      #   Source: Robotiq_Grippers, 1.8.4.4844, Robotiq Inc.
      #   Type: Gripper
      $ 2003 "Gripper Close (1)"
      if not(gripper_connected[0]):
        popup("Gripper 1 must be connected to run this program.", "No connection", False, True, True)
      end
      if not(rq_is_gripper_activated("1")):
        popup("Gripper 1 is not activated. Go to Installation tab > Gripper to activate it and run the program again.", "Not activated", False, True, True)
      end
      rq_set_pos_spd_for(255, 204, 255, "1")
      rq_wait_pos_spe_for_request(255, 204, 255, "1")
      rq_go_to("1")
      rq_wait("1")
      # end: URCap Program Node
      $ 2010 "Decap"
      $ 2011 "Action_Info≔'decapping'"
      global Action_Info="decapping"
      $ 2012 "Set GRP_3F_Enable=On"
      set_standard_digital_out(4, True)
      $ 2013 "Set GRP_3F_Decap=On"
      set_standard_digital_out(3, True)
      $ 2014 "Force"
      sleep(0.02)
      zero_ftsensor()
      force_mode(p[0.0,0.0,0.0,0.0,0.0,0.0], [0, 0, 1, 0, 0, 0], [0.0, 0.0, 1.0, 0.0, 0.0, 0.0], 2, [0.1, 0.1, 0.001, 0.3490658503988659, 0.3490658503988659, 0.3490658503988659])
      $ 2015 "check_decapping(offset=0.015, timeout=10, abort=CMD_Hold)" "noBreak"
      check_decapping(offset=0.015, timeout=10, abort=CMD_Hold)
      end_force_mode()
      stopl(5.0)
      $ 2016 "Set GRP_3F_Decap=Off"
      set_standard_digital_out(3, False)
      $ 2017 "Set GRP_3F_Enable=Off"
      set_standard_digital_out(4, False)
      $ 2018 "MoveL"
      $ 2019 "Waypoint_50" "breakAfter"
      movel(Waypoint_50_p, a=0.5, v=0.1, r=0.05)
      $ 2020 "MoveJ"
      $ 2021 "cap_dump" "breakAfter"
      movej(get_inverse_kin(cap_dump_p, qnear=cap_dump_q), a=0.5235987755982988, v=0.4363323129985824)
      # begin: URCap Program Node
      #   Source: Robotiq_Grippers, 1.8.4.4844, Robotiq Inc.
      #   Type: Gripper
      $ 2022 "Gripper Open (1)"
      if not(gripper_connected[0]):
        popup("Gripper 1 must be connected to run this program.", "No connection", False, True, True)
      end
      if not(rq_is_gripper_activated("1")):
        popup("Gripper 1 is not activated. Go to Installation tab > Gripper to activate it and run the program again.", "Not activated", False, True, True)
      end
      rq_set_pos_spd_for(0, 204, 255, "1")
      rq_wait_pos_spe_for_request(0, 204, 255, "1")
      rq_go_to("1")
      rq_wait("1")
      # end: URCap Program Node
      $ 2023 "MoveJ"
      $ 2024 "Waypoint_51" "breakAfter"
      movej(get_inverse_kin(Waypoint_51_p, qnear=Waypoint_51_q), a=0.5235987755982988, v=0.4363323129985824, r=0.036)
    elif (33 == switch_1):
      $ 2025 "Case 33"
      $ 2026 "Shake and liquid transfer"
      $ 2027 "MoveL"
      $ 2028 "Vial_liq_above" "breakAfter"
      movel(Vial_liq_above_p, a=0.5, v=0.1)
      $ 2029 "Vial_liq_pick_1" "breakAfter"
      movel(Vial_liq_pick_1_p, a=0.5, v=0.1)
      $ 2030 "Vial_liq_pick_2" "breakAfter"
      movel(Vial_liq_pick_2_p, a=0.5, v=0.1)
      # begin: URCap Program Node
      #   Source: Robotiq_Grippers, 1.8.4.4844, Robotiq Inc.
      #   Type: Gripper
      $ 2031 "Gripper Close (1)"
      if not(gripper_connected[0]):
        popup("Gripper 1 must be connected to run this program.", "No connection", False, True, True)
      end
      if not(rq_is_gripper_activated("1")):
        popup("Gripper 1 is not activated. Go to Installation tab > Gripper to activate it and run the program again.", "Not activated", False, True, True)
      end
      rq_set_pos_spd_for(255, 82, 71, "1")
      rq_wait_pos_spe_for_request(255, 82, 71, "1")
      rq_go_to("1")
      rq_wait("1")
      # end: URCap Program Node
      $ 2032 "Wait: 1.0"
      sleep(1.0)
      $ 2033 "Set GRP_3F_Open=On"
      set_standard_digital_out(5, True)
      $ 2034 "Wait: 0.5"
      sleep(0.5)
      $ 2035 "Vial_liq_above" "breakAfter"
      movel(Vial_liq_above_p, a=0.3, v=0.05, r=0.05)
      $ 2036 "MoveL"
      $ 2037 "Liquid_midway" "breakAfter"
      movel(Liquid_midway_p, a=0.5, v=0.1)
      $ 2038 "Loop 3 times"
      Loop_1 = 0
      while (Loop_1 < 3):
        $ 2039 "shake_1" "breakAfter"
        movel(shake_1_p, a=2.0, v=0.5)
        $ 2040 "shake_2" "breakAfter"
        movel(shake_2_p, a=2.0, v=0.5)
        Loop_1 = Loop_1 + 1
      end
      $ 2041 "drop_above_1" "breakAfter"
      movel(drop_above_1_p, a=0.5, v=0.1)
      $ 2042 "drop_above_2" "breakAfter"
      movel(drop_above_2_p, a=0.5, v=0.1)
      $ 2043 "liq_tran_1" "breakAfter"
      movel(liq_tran_1_p, a=0.5, v=0.05, r=0.008)
      $ 2044 "Wait: 1.0"
      sleep(1.0)
      $ 2045 "drop_above_2" "breakAfter"
      movel(drop_above_2_p, a=0.5, v=0.1)
      $ 2046 "Waypoint_21" "breakAfter"
      movel(Waypoint_21_p, a=0.5, v=0.1)
      $ 2047 "liq_tran_2" "breakAfter"
      movel(liq_tran_2_p, a=0.5, v=0.05)
      $ 2048 "Wait: 1.0"
      sleep(1.0)
      $ 2049 "drop_above_2" "breakAfter"
      movel(drop_above_2_p, a=0.5, v=0.1)
      $ 2050 "drop_above_1" "breakAfter"
      movel(drop_above_1_p, a=0.5, v=0.1)
      $ 2051 "Liquid_midway" "breakAfter"
      movel(Liquid_midway_p, a=0.5, v=0.1)
      $ 2052 "MoveL"
      $ 2053 "Vial_drop_above" "breakAfter"
      movel(Vial_drop_above_p, a=0.5, v=0.1)
      $ 2054 "Vial_liq_drop" "breakAfter"
      movel(Vial_liq_drop_p, a=0.5, v=0.1)
      # begin: URCap Program Node
      #   Source: Robotiq_Grippers, 1.8.4.4844, Robotiq Inc.
      #   Type: Gripper
      $ 2055 "Gripper Open (1)"
      if not(gripper_connected[0]):
        popup("Gripper 1 must be connected to run this program.", "No connection", False, True, True)
      end
      if not(rq_is_gripper_activated("1")):
        popup("Gripper 1 is not activated. Go to Installation tab > Gripper to activate it and run the program again.", "Not activated", False, True, True)
      end
      rq_set_pos_spd_for(0, 82, 71, "1")
      rq_wait_pos_spe_for_request(0, 82, 71, "1")
      rq_go_to("1")
      rq_wait("1")
      # end: URCap Program Node
      $ 2056 "Vial_drop_above" "breakAfter"
      movel(Vial_drop_above_p, a=0.5, v=0.1)
    elif (34 == switch_1):
      $ 2057 "Case 34"
      $ 2058 "Home (Safe)"
      movej([-1.2302089344500047, -1.2969853503591224, -1.875639182904262, -1.539621866126728, 1.5731943360401213, -2.80099559440227], a=1.3962634015954636, v=1.0471975511965976)
      $ 2059 "MoveJ"
      $ 2060 "Waypoint_9" "breakAfter"
      movej(get_inverse_kin(Waypoint_9_p, qnear=Waypoint_9_q), a=0.5235987755982988, v=0.4363323129985824)
      $ 2061 "MoveL"
      $ 2062 "Waypoint_10" "breakAfter"
      movel(Waypoint_10_p, a=0.5, v=0.1)
      # begin: URCap Program Node
      #   Source: Robotiq_Grippers, 1.8.4.4844, Robotiq Inc.
      #   Type: Gripper
      $ 2063 "Gripper Close (1)"
      if not(gripper_connected[0]):
        popup("Gripper 1 must be connected to run this program.", "No connection", False, True, True)
      end
      if not(rq_is_gripper_activated("1")):
        popup("Gripper 1 is not activated. Go to Installation tab > Gripper to activate it and run the program again.", "Not activated", False, True, True)
      end
      rq_set_pos_spd_for(255, 82, 71, "1")
      rq_wait_pos_spe_for_request(255, 82, 71, "1")
      rq_go_to("1")
      rq_wait("1")
      # end: URCap Program Node
      $ 2064 "Wait: 1.0"
      sleep(1.0)
      $ 2065 "MoveL"
      $ 2066 "Waypoint_11" "breakAfter"
      movel(Waypoint_11_p, a=0.5, v=0.1, r=0.05)
      $ 2067 "MoveJ"
      $ 2068 "Waypoint_7" "breakAfter"
      movej(get_inverse_kin(Waypoint_7_p, qnear=Waypoint_7_q), a=0.5235987755982988, v=0.4363323129985824, r=0.05)
      $ 2069 "MoveL"
      $ 2070 "Waypoint_8" "breakAfter"
      movel(Waypoint_8_p, a=0.5, v=0.1)
      # begin: URCap Program Node
      #   Source: Robotiq_Grippers, 1.8.4.4844, Robotiq Inc.
      #   Type: Gripper
      $ 2071 "Gripper Open (1)"
      if not(gripper_connected[0]):
        popup("Gripper 1 must be connected to run this program.", "No connection", False, True, True)
      end
      if not(rq_is_gripper_activated("1")):
        popup("Gripper 1 is not activated. Go to Installation tab > Gripper to activate it and run the program again.", "Not activated", False, True, True)
      end
      rq_set_pos_spd_for(0, 82, 71, "1")
      rq_wait_pos_spe_for_request(0, 82, 71, "1")
      rq_go_to("1")
      rq_wait("1")
      # end: URCap Program Node
      $ 2072 "MoveJ"
      $ 2073 "Waypoint_7" "breakAfter"
      movej(get_inverse_kin(Waypoint_7_p, qnear=Waypoint_7_q), a=0.5235987755982988, v=0.4363323129985824)
      $ 2074 "Home (Safe)"
      movej([-1.2302089344500047, -1.2969853503591224, -1.875639182904262, -1.539621866126728, 1.5731943360401213, -2.80099559440227], a=1.3962634015954636, v=1.0471975511965976)
    elif (35 == switch_1):
      $ 2091 "Case 35"
      $ 2092 "Pick the powder container"
      $ 2093 "Wait: 1.0"
      sleep(1.0)
      $ 2094 "MoveJ"
      $ 2095 "Container_midwa" "breakAfter"
      movej(get_inverse_kin(Container_midwa_p, qnear=Container_midwa_q), a=1.3962634015954636, v=1.0471975511965976, r=0.05)
      $ 2096 "Container_capt" "breakAfter"
      movej(get_inverse_kin(Container_capt_p, qnear=Container_capt_q), a=1.3962634015954636, v=1.0471975511965976)
      # begin: URCap Program Node
      #   Source: SensoPart VISOR Robotic, 2.0.0, SensoPart Industriesensorik GmbH
      #   Type: VISOR Robotic App
      $ 2097 "VISOR Easy Pick"
      def visorFuncEasyPick_e3134b():
        # begin: URCap Program Node
        #   Source: SensoPart VISOR Robotic, 2.0.0, SensoPart Industriesensorik GmbH
        #   Type: Easy Pick Setup
        $ 2098 "# 1 Setup" "noBreak"
        local easyPickVisorId = 1
        local easyPickArmMounted = True
        local easyPickSetJob = True
        local easyPickJobName = "Container_S"
        local easyPickAtImgAcq = False
        local easyPickImgAcqPose = p[-0.5104,0.4173,0.4641,0.0000,-0.0000,-2.8962]
        # end: URCap Program Node
        # begin: URCap Program Node
        #   Source: SensoPart VISOR Robotic, 2.0.0, SensoPart Industriesensorik GmbH
        #   Type: Process
        $ 2099 "Process" "noBreak"
        local easyPickObjTaken = False
        local easyPickTrigger = False
        local easyPickPoseIdx = 0
        local easyPickPose = p[0,0,0,0,0,0]
        def easyPickFuncTrigger(visorId, setJob, jobName, arm):
        if (setJob):
          visor_changeJob(visorId, jobName, 6000)
        end
        if (arm):
          visor_trigger(visorId, 6000, "arm")
        else:
          visor_trigger(visorId, 6000)
        end
        global easyPickParts=visor_partsFound(visorId)
        visor_easyPickUpdate(visorId, "parts", visor_partsFound(visorId))
        return visor_getPose3d(visorId, 0)
      end
      while (not easyPickObjTaken):
        easyPickTrigger = (easyPickCount >= visor_partsFound(easyPickVisorId)) or (easyPickCount > 9) or (not visor_easyPickCheckIdent("70ff7e", easyPickVisorId))
        if (easyPickTrigger):
          easyPickCount = 0
        end
        easyPickPoseIdx = easyPickCount
        easyPickPose = visor_getPose3d(easyPickVisorId, easyPickPoseIdx)
        visor_easyPickUpdate(easyPickVisorId, "counter", easyPickPoseIdx)
        # begin: URCap Program Node
        #   Source: SensoPart VISOR Robotic, 2.0.0, SensoPart Industriesensorik GmbH
        #   Type: Image Acquisition Pose
        $ 2100 "Image Acquisition Pose" "noBreak"
        if (easyPickTrigger):
          if (not easyPickAtImgAcq):
            movej(pose_trans(easyPickImgAcqPose,p[0.0000,0.0000,-0.0000,0.0000,0.0000,0.0000]),a=1.3963,v=1.0472,t=0.000000,r=0.000000)
            easyPickAtImgAcq = True
          end
          easyPickPose = easyPickFuncTrigger(easyPickVisorId, easyPickSetJob, easyPickJobName, easyPickArmMounted)
        end
        # end: URCap Program Node
        # begin: URCap Program Node
        #   Source: SensoPart VISOR Robotic, 2.0.0, SensoPart Industriesensorik GmbH
        #   Type: Object Detected
        $ 2101 "Object Detected" "noBreak"
        if (visor_partsFound(easyPickVisorId) > 0):
          $ 2102 "Open Gripper" "noBreak"
          # begin: URCap Program Node
          #   Source: Robotiq_Grippers, 1.8.4.4844, Robotiq Inc.
          #   Type: Gripper
          $ 2103 "Gripper Open (1)" "noBreak"
          if not(gripper_connected[0]):
            popup("Gripper 1 must be connected to run this program.", "No connection", False, True, True)
          end
          if not(rq_is_gripper_activated("1")):
            popup("Gripper 1 is not activated. Go to Installation tab > Gripper to activate it and run the program again.", "Not activated", False, True, True)
          end
          rq_set_pos_spd_for(0, 107, 77, "1")
          rq_wait_pos_spe_for_request(0, 107, 77, "1")
          rq_go_to("1")
          rq_wait("1")
          # end: URCap Program Node
          $ 2104 "MoveJ" "noBreak"
          $ 2105 "Waypoint_13" "noBreak"
          movej(get_inverse_kin(Waypoint_13_p, qnear=Waypoint_13_q), a=1.3962634015954636, v=1.0471975511965976)
          # begin: URCap Program Node
          #   Source: SensoPart VISOR Robotic, 2.0.0, SensoPart Industriesensorik GmbH
          #   Type: Approach Pose
          $ 2106 "Approach Pose" "noBreak"
          movej(pose_trans(easyPickPose,p[0.0000,0.0000,0.0500,0.0000,0.0000,0.0000]),a=1.3963,v=1.0472,t=0.000000,r=0.000000)
          # end: URCap Program Node
          # begin: URCap Program Node
          #   Source: SensoPart VISOR Robotic, 2.0.0, SensoPart Industriesensorik GmbH
          #   Type: Target Pose
          $ 2107 "Target Pose" "noBreak"
          movel(pose_trans(easyPickPose,p[0.0000,0.0000,-0.0000,0.0000,0.0000,0.0000]),a=0.5000,v=0.2500,t=0.000000,r=0.000000)
          # end: URCap Program Node
          $ 2108 "Close Gripper" "noBreak"
          # begin: URCap Program Node
          #   Source: Robotiq_Grippers, 1.8.4.4844, Robotiq Inc.
          #   Type: Gripper
          $ 2109 "Gripper Close (1)" "noBreak"
          if not(gripper_connected[0]):
            popup("Gripper 1 must be connected to run this program.", "No connection", False, True, True)
          end
          if not(rq_is_gripper_activated("1")):
            popup("Gripper 1 is not activated. Go to Installation tab > Gripper to activate it and run the program again.", "Not activated", False, True, True)
          end
          rq_set_pos_spd_for(255, 107, 77, "1")
          rq_wait_pos_spe_for_request(255, 107, 77, "1")
          rq_go_to("1")
          rq_wait("1")
          # end: URCap Program Node
          # begin: URCap Program Node
          #   Source: SensoPart VISOR Robotic, 2.0.0, SensoPart Industriesensorik GmbH
          #   Type: Exit Pose
          $ 2110 "Exit Pose" "noBreak"
          movel(pose_trans(easyPickPose,p[0.0000,0.0000,0.0500,0.0000,0.0000,0.0000]),a=0.5000,v=0.2500,t=0.000000,r=0.000000)
          # end: URCap Program Node
          easyPickObjTaken = True
        end
        # end: URCap Program Node
        # begin: URCap Program Node
        #   Source: SensoPart VISOR Robotic, 2.0.0, SensoPart Industriesensorik GmbH
        #   Type: No Object Detected
        $ 2111 "No Object Detected" "noBreak"
        if (visor_partsFound(easyPickVisorId) < 1):
          easyPickNoObj = easyPickNoObj + 1
          if (easyPickNoObj > 5):
            global easyPickNoObj=0
            halt
          end
          $ 2112 "Popup: No Container detected" "noBreak"
          popup("No Container detected", "Message", False, False, blocking=True)
          else:
          global easyPickNoObj=0
        end
        # end: URCap Program Node
      end
      easyPickCount = easyPickCount + 1
      visor_easyPickUpdate(easyPickVisorId, "counter", easyPickCount)
      visor_easyPickSetIdent("70ff7e", easyPickVisorId)
      # end: URCap Program Node
    end
    visorFuncEasyPick_e3134b()
    # end: URCap Program Node
    $ 2113 "MoveJ"
    $ 2114 "Cont_midwa_1" "breakAfter"
    movej(get_inverse_kin(Cont_midwa_1_p, qnear=Cont_midwa_1_q), a=1.3962634015954636, v=1.0471975511965976, r=0.05)
    $ 2115 "Cont_midw_2" "breakAfter"
    movej(get_inverse_kin(Cont_midw_2_p, qnear=Cont_midw_2_q), a=1.3962634015954636, v=1.0471975511965976, r=0.05)
    $ 2116 "MoveJ"
    $ 2117 "Waypoint_14" "breakAfter"
    movej(get_inverse_kin(Waypoint_14_p, qnear=Waypoint_14_q), a=1.3962634015954636, v=1.0471975511965976)
    $ 2118 "Cont_midway_3" "breakAfter"
    movej(get_inverse_kin(Cont_midway_3_p, qnear=Cont_midway_3_q), a=1.3962634015954636, v=1.0471975511965976)
    $ 2119 "Waypoint_43" "breakAfter"
    movej(get_inverse_kin(Waypoint_43_p, qnear=Waypoint_43_q), a=1.3962634015954636, v=1.0471975511965976)
    $ 2120 "MoveL"
    $ 2121 "Waypoint_27" "breakAfter"
    movel(Waypoint_27_p, a=1.2, v=0.25)
    $ 2122 "Waypoint_2" "breakAfter"
    movel(Waypoint_2_p, a=0.3, v=0.05)
    # begin: URCap Program Node
    #   Source: Robotiq_Grippers, 1.8.4.4844, Robotiq Inc.
    #   Type: Gripper
    $ 2123 "Gripper Open (1)"
    if not(gripper_connected[0]):
      popup("Gripper 1 must be connected to run this program.", "No connection", False, True, True)
    end
    if not(rq_is_gripper_activated("1")):
      popup("Gripper 1 is not activated. Go to Installation tab > Gripper to activate it and run the program again.", "Not activated", False, True, True)
    end
    rq_set_pos_spd_for(0, 255, 255, "1")
    rq_wait_pos_spe_for_request(0, 255, 255, "1")
    rq_go_to("1")
    rq_wait("1")
    # end: URCap Program Node
    $ 2124 "MoveL"
    $ 2125 "Waypoint_27" "breakAfter"
    movel(Waypoint_27_p, a=1.2, v=0.25)
    $ 2126 "Waypoint_39" "breakAfter"
    movel(Waypoint_39_p, a=1.2, v=0.25)
    $ 2127 "Home (Safe)"
    movej([-1.2302089344500047, -1.2969853503591224, -1.875639182904262, -1.539621866126728, 1.5731943360401213, -2.80099559440227], a=1.3962634015954636, v=1.0471975511965976)
    # begin: URCap Program Node
    #   Source: SensoPart VISOR Robotic, 2.0.0, SensoPart Industriesensorik GmbH
    #   Type: VISOR Robotic App
    $ 2128 "VISOR Easy Pick"
    def visorFuncEasyPick_ffc504():
      # begin: URCap Program Node
      #   Source: SensoPart VISOR Robotic, 2.0.0, SensoPart Industriesensorik GmbH
      #   Type: Easy Pick Setup
      $ 2129 "# 1 Setup" "noBreak"
      local easyPickVisorId = 1
      local easyPickArmMounted = True
      local easyPickSetJob = True
      local easyPickJobName = "Target_container"
      local easyPickAtImgAcq = False
      local easyPickImgAcqPose = p[-0.6180,0.3719,0.4116,-0.0000,-0.0000,-2.8962]
      # end: URCap Program Node
      # begin: URCap Program Node
      #   Source: SensoPart VISOR Robotic, 2.0.0, SensoPart Industriesensorik GmbH
      #   Type: Process
      $ 2130 "Process" "noBreak"
      local easyPickObjTaken = False
      local easyPickTrigger = False
      local easyPickPoseIdx = 0
      local easyPickPose = p[0,0,0,0,0,0]
      def easyPickFuncTrigger(visorId, setJob, jobName, arm):
      if (setJob):
        visor_changeJob(visorId, jobName, 6000)
      end
      if (arm):
        visor_trigger(visorId, 6000, "arm")
      else:
        visor_trigger(visorId, 6000)
      end
      global easyPickParts_2=visor_partsFound(visorId)
      visor_easyPickUpdate(visorId, "parts", visor_partsFound(visorId))
      return visor_getPose3d(visorId, 0)
    end
    while (not easyPickObjTaken):
      easyPickTrigger = (easyPickCount_2 >= visor_partsFound(easyPickVisorId)) or (easyPickCount_2 > 9) or (not visor_easyPickCheckIdent("9ee82b", easyPickVisorId))
      if (easyPickTrigger):
        easyPickCount_2 = 0
      end
      easyPickPoseIdx = easyPickCount_2
      easyPickPose = visor_getPose3d(easyPickVisorId, easyPickPoseIdx)
      visor_easyPickUpdate(easyPickVisorId, "counter", easyPickPoseIdx)
      # begin: URCap Program Node
      #   Source: SensoPart VISOR Robotic, 2.0.0, SensoPart Industriesensorik GmbH
      #   Type: Image Acquisition Pose
      $ 2131 "Image Acquisition Pose" "noBreak"
      if (easyPickTrigger):
        if (not easyPickAtImgAcq):
          movej(pose_trans(easyPickImgAcqPose,p[0.0000,0.0000,-0.0000,0.0000,0.0000,0.0000]),a=1.3963,v=1.0472,t=0.000000,r=0.000000)
          easyPickAtImgAcq = True
        end
        easyPickPose = easyPickFuncTrigger(easyPickVisorId, easyPickSetJob, easyPickJobName, easyPickArmMounted)
      end
      # end: URCap Program Node
      # begin: URCap Program Node
      #   Source: SensoPart VISOR Robotic, 2.0.0, SensoPart Industriesensorik GmbH
      #   Type: Object Detected
      $ 2132 "Object Detected" "noBreak"
      if (visor_partsFound(easyPickVisorId) > 0):
        $ 2133 "Open Gripper" "noBreak"
        # begin: URCap Program Node
        #   Source: Robotiq_Grippers, 1.8.4.4844, Robotiq Inc.
        #   Type: Gripper
        $ 2134 "Gripper Open (1)" "noBreak"
        if not(gripper_connected[0]):
          popup("Gripper 1 must be connected to run this program.", "No connection", False, True, True)
        end
        if not(rq_is_gripper_activated("1")):
          popup("Gripper 1 is not activated. Go to Installation tab > Gripper to activate it and run the program again.", "Not activated", False, True, True)
        end
        rq_set_pos_spd_for(0, 107, 77, "1")
        rq_wait_pos_spe_for_request(0, 107, 77, "1")
        rq_go_to("1")
        rq_wait("1")
        # end: URCap Program Node
        # begin: URCap Program Node
        #   Source: SensoPart VISOR Robotic, 2.0.0, SensoPart Industriesensorik GmbH
        #   Type: Approach Pose
        $ 2135 "Approach Pose" "noBreak"
        movej(pose_trans(easyPickPose,p[0.0000,0.0000,0.0500,0.0000,0.0000,0.0000]),a=1.3963,v=1.0472,t=0.000000,r=0.000000)
        # end: URCap Program Node
        # begin: URCap Program Node
        #   Source: SensoPart VISOR Robotic, 2.0.0, SensoPart Industriesensorik GmbH
        #   Type: Target Pose
        $ 2136 "Target Pose" "noBreak"
        movel(pose_trans(easyPickPose,p[0.0000,0.0000,-0.0000,0.0000,0.0000,0.0000]),a=0.5000,v=0.2500,t=0.000000,r=0.000000)
        # end: URCap Program Node
        $ 2137 "Close Gripper" "noBreak"
        # begin: URCap Program Node
        #   Source: Robotiq_Grippers, 1.8.4.4844, Robotiq Inc.
        #   Type: Gripper
        $ 2138 "Gripper Close (1)" "noBreak"
        if not(gripper_connected[0]):
          popup("Gripper 1 must be connected to run this program.", "No connection", False, True, True)
        end
        if not(rq_is_gripper_activated("1")):
          popup("Gripper 1 is not activated. Go to Installation tab > Gripper to activate it and run the program again.", "Not activated", False, True, True)
        end
        rq_set_pos_spd_for(255, 107, 77, "1")
        rq_wait_pos_spe_for_request(255, 107, 77, "1")
        rq_go_to("1")
        rq_wait("1")
        # end: URCap Program Node
        # begin: URCap Program Node
        #   Source: SensoPart VISOR Robotic, 2.0.0, SensoPart Industriesensorik GmbH
        #   Type: Exit Pose
        $ 2139 "Exit Pose" "noBreak"
        movel(pose_trans(easyPickPose,p[0.0000,0.0000,0.0500,0.0000,0.0000,0.0000]),a=0.5000,v=0.2500,t=0.000000,r=0.000000)
        # end: URCap Program Node
        easyPickObjTaken = True
      end
      # end: URCap Program Node
      # begin: URCap Program Node
      #   Source: SensoPart VISOR Robotic, 2.0.0, SensoPart Industriesensorik GmbH
      #   Type: No Object Detected
      $ 2140 "No Object Detected" "noBreak"
      if (visor_partsFound(easyPickVisorId) < 1):
        easyPickNoObj_2 = easyPickNoObj_2 + 1
        if (easyPickNoObj_2 > 5):
          global easyPickNoObj_2=0
          halt
        end
        $ 2141 "Popup: No target container is detected" "noBreak"
        popup("No target container is detected", "Message", False, False, blocking=True)
        else:
        global easyPickNoObj_2=0
      end
      # end: URCap Program Node
    end
    easyPickCount_2 = easyPickCount_2 + 1
    visor_easyPickUpdate(easyPickVisorId, "counter", easyPickCount_2)
    visor_easyPickSetIdent("9ee82b", easyPickVisorId)
    # end: URCap Program Node
  end
  visorFuncEasyPick_ffc504()
  # end: URCap Program Node
  $ 2142 "MoveJ"
  $ 2143 "Waypoint_5" "breakAfter"
  movej(get_inverse_kin(Waypoint_5_p, qnear=Waypoint_5_q), a=1.3962634015954636, v=1.0471975511965976)
  $ 2144 "Waypoint_3" "breakAfter"
  movej(get_inverse_kin(Waypoint_3_p, qnear=Waypoint_3_q), a=1.3962634015954636, v=1.0471975511965976)
  $ 2145 "Set GRP_3F_Open=On"
  set_standard_digital_out(5, True)
  $ 2146 "MoveL"
  $ 2147 "Waypoint_4" "breakAfter"
  movel(Waypoint_4_p, a=1.2, v=0.25)
  $ 2148 "Waypoint_15" "breakAfter"
  movel(Waypoint_15_p, a=0.3, v=0.05)
  $ 2149 "Set GRP_3F_Open=Off"
  set_standard_digital_out(5, False)
  $ 2150 "Wait: 0.5"
  sleep(0.5)
  # begin: URCap Program Node
  #   Source: Robotiq_Grippers, 1.8.4.4844, Robotiq Inc.
  #   Type: Gripper
  $ 2151 "Gripper Open (1)"
  if not(gripper_connected[0]):
    popup("Gripper 1 must be connected to run this program.", "No connection", False, True, True)
  end
  if not(rq_is_gripper_activated("1")):
    popup("Gripper 1 is not activated. Go to Installation tab > Gripper to activate it and run the program again.", "Not activated", False, True, True)
  end
  rq_set_pos_spd_for(0, 127, 71, "1")
  rq_wait_pos_spe_for_request(0, 127, 71, "1")
  rq_go_to("1")
  rq_wait("1")
  # end: URCap Program Node
  $ 2152 "MoveL"
  $ 2153 "Waypoint_16" "breakAfter"
  movel(Waypoint_16_p, a=1.2, v=0.25)
  $ 2154 "Home (Safe)"
  movej([-1.2302089344500047, -1.2969853503591224, -1.875639182904262, -1.539621866126728, 1.5731943360401213, -2.80099559440227], a=1.3962634015954636, v=1.0471975511965976)
  elif (36 == switch_1):
    $ 2155 "Case 36"
    $ 2156 "MoveJ"
    $ 2157 "Waypoint_23" "breakAfter"
    movej(get_inverse_kin(Waypoint_23_p, qnear=Waypoint_23_q), a=1.3962634015954636, v=1.0471975511965976)
    $ 2158 "MoveL"
    $ 2159 "Waypoint_24" "breakAfter"
    movel(Waypoint_24_p, a=1.2, v=0.25)
    # begin: URCap Program Node
    #   Source: Robotiq_Grippers, 1.8.4.4844, Robotiq Inc.
    #   Type: Gripper
    $ 2160 "Gripper Close (1)"
    if not(gripper_connected[0]):
      popup("Gripper 1 must be connected to run this program.", "No connection", False, True, True)
    end
    if not(rq_is_gripper_activated("1")):
      popup("Gripper 1 is not activated. Go to Installation tab > Gripper to activate it and run the program again.", "Not activated", False, True, True)
    end
    rq_set_pos_spd_for(255, 127, 127, "1")
    rq_wait_pos_spe_for_request(255, 127, 127, "1")
    rq_go_to("1")
    rq_wait("1")
    # end: URCap Program Node
    $ 2161 "Decap"
    $ 2162 "Action_Info≔'decapping'"
    global Action_Info="decapping"
    $ 2163 "Set GRP_3F_Enable=On"
    set_standard_digital_out(4, True)
    $ 2164 "Set GRP_3F_Decap=On"
    set_standard_digital_out(3, True)
    $ 2165 "Force"
    sleep(0.02)
    zero_ftsensor()
    force_mode(p[0.0,0.0,0.0,0.0,0.0,0.0], [0, 0, 1, 0, 0, 0], [0.0, 0.0, 1.0, 0.0, 0.0, 0.0], 2, [0.1, 0.1, 0.001, 0.3490658503988659, 0.3490658503988659, 0.3490658503988659])
    $ 2166 "check_decapping(offset=0.08, timeout=16, abort=CMD_Hold)" "noBreak"
    check_decapping(offset=0.08, timeout=16, abort=CMD_Hold)
    end_force_mode()
    stopl(5.0)
    $ 2167 "Set GRP_3F_Decap=Off"
    set_standard_digital_out(3, False)
    $ 2168 "Set GRP_3F_Enable=Off"
    set_standard_digital_out(4, False)
    $ 2169 "MoveL"
    $ 2170 "Waypoint_17" "breakAfter"
    movel(Waypoint_17_p, a=1.2, v=0.25)
    $ 2171 "Waypoint_22" "breakAfter"
    movel(Waypoint_22_p, a=1.2, v=0.25)
    $ 2172 "Waypoint_25" "breakAfter"
    movel(Waypoint_25_p, a=1.2, v=0.25)
    # begin: URCap Program Node
    #   Source: Robotiq_Grippers, 1.8.4.4844, Robotiq Inc.
    #   Type: Gripper
    $ 2173 "Gripper Open (1)"
    if not(gripper_connected[0]):
      popup("Gripper 1 must be connected to run this program.", "No connection", False, True, True)
    end
    if not(rq_is_gripper_activated("1")):
      popup("Gripper 1 is not activated. Go to Installation tab > Gripper to activate it and run the program again.", "Not activated", False, True, True)
    end
    rq_set_pos_spd_for(0, 107, 77, "1")
    rq_wait_pos_spe_for_request(0, 107, 77, "1")
    rq_go_to("1")
    rq_wait("1")
    # end: URCap Program Node
    $ 2174 "MoveL"
    $ 2175 "Waypoint_26" "breakAfter"
    movel(Waypoint_26_p, a=1.2, v=0.25)
    $ 2176 "MoveL"
    $ 2177 "Waypoint_30" "breakAfter"
    movel(Waypoint_30_p, a=1.2, v=0.25)
    $ 2178 "Waypoint_28" "breakAfter"
    movel(Waypoint_28_p, a=1.2, v=0.25)
    # begin: URCap Program Node
    #   Source: Robotiq_Grippers, 1.8.4.4844, Robotiq Inc.
    #   Type: Gripper
    $ 2179 "Gripper Close (1)"
    if not(gripper_connected[0]):
      popup("Gripper 1 must be connected to run this program.", "No connection", False, True, True)
    end
    if not(rq_is_gripper_activated("1")):
      popup("Gripper 1 is not activated. Go to Installation tab > Gripper to activate it and run the program again.", "Not activated", False, True, True)
    end
    rq_set_pos_spd_for(255, 107, 77, "1")
    rq_wait_pos_spe_for_request(255, 107, 77, "1")
    rq_go_to("1")
    rq_wait("1")
    # end: URCap Program Node
    $ 2180 "Wait: 0.5"
    sleep(0.5)
    $ 2181 "Set GRP_3F_Open=On"
    set_standard_digital_out(5, True)
    $ 2182 "MoveL"
    $ 2183 "Waypoint_29" "breakAfter"
    movel(Waypoint_29_p, a=1.2, v=0.25)
    $ 2184 "MoveJ"
    $ 2185 "Waypoint_31" "breakAfter"
    movej(get_inverse_kin(Waypoint_31_p, qnear=Waypoint_31_q), a=1.3962634015954636, v=1.0471975511965976)
    # begin: URCap Program Node
    #   Source: SensoPart VISOR Robotic, 2.0.0, SensoPart Industriesensorik GmbH
    #   Type: VISOR Robotic App
    $ 2186 "VISOR Easy Pick"
    def visorFuncEasyPick_7a8a4a():
      # begin: URCap Program Node
      #   Source: SensoPart VISOR Robotic, 2.0.0, SensoPart Industriesensorik GmbH
      #   Type: Easy Pick Setup
      $ 2187 "# 1 Setup" "noBreak"
      local easyPickVisorId = 1
      local easyPickArmMounted = True
      local easyPickSetJob = True
      local easyPickJobName = "Weigh_scale"
      local easyPickAtImgAcq = False
      local easyPickImgAcqPose = p[-0.6121,0.0166,0.5300,0.0440,-0.0067,-1.6589]
      # end: URCap Program Node
      # begin: URCap Program Node
      #   Source: SensoPart VISOR Robotic, 2.0.0, SensoPart Industriesensorik GmbH
      #   Type: Process
      $ 2188 "Process" "noBreak"
      local easyPickObjTaken = False
      local easyPickTrigger = False
      local easyPickPoseIdx = 0
      local easyPickPose = p[0,0,0,0,0,0]
      def easyPickFuncTrigger(visorId, setJob, jobName, arm):
      if (setJob):
        visor_changeJob(visorId, jobName, 6000)
      end
      if (arm):
        visor_trigger(visorId, 6000, "arm")
      else:
        visor_trigger(visorId, 6000)
      end
      global easyPickParts_1=visor_partsFound(visorId)
      visor_easyPickUpdate(visorId, "parts", visor_partsFound(visorId))
      return visor_getPose3d(visorId, 0)
    end
    while (not easyPickObjTaken):
      easyPickTrigger = (easyPickCount_1 >= visor_partsFound(easyPickVisorId)) or (easyPickCount_1 > 9) or (not visor_easyPickCheckIdent("425780", easyPickVisorId))
      if (easyPickTrigger):
        easyPickCount_1 = 0
      end
      easyPickPoseIdx = easyPickCount_1
      easyPickPose = visor_getPose3d(easyPickVisorId, easyPickPoseIdx)
      visor_easyPickUpdate(easyPickVisorId, "counter", easyPickPoseIdx)
      # begin: URCap Program Node
      #   Source: SensoPart VISOR Robotic, 2.0.0, SensoPart Industriesensorik GmbH
      #   Type: Image Acquisition Pose
      $ 2189 "Image Acquisition Pose" "noBreak"
      if (easyPickTrigger):
        if (not easyPickAtImgAcq):
          movej(pose_trans(easyPickImgAcqPose,p[0.0000,0.0000,-0.0000,0.0000,0.0000,0.0000]),a=1.3963,v=1.0472,t=0.000000,r=0.000000)
          easyPickAtImgAcq = True
        end
        easyPickPose = easyPickFuncTrigger(easyPickVisorId, easyPickSetJob, easyPickJobName, easyPickArmMounted)
      end
      # end: URCap Program Node
      # begin: URCap Program Node
      #   Source: SensoPart VISOR Robotic, 2.0.0, SensoPart Industriesensorik GmbH
      #   Type: Object Detected
      $ 2190 "Object Detected" "noBreak"
      if (visor_partsFound(easyPickVisorId) > 0):
        $ 2191 "Open Gripper" "noBreak"
        $ 2192 "Wait: 0.5" "noBreak"
        sleep(0.5)
        # begin: URCap Program Node
        #   Source: SensoPart VISOR Robotic, 2.0.0, SensoPart Industriesensorik GmbH
        #   Type: Approach Pose
        $ 2193 "Approach Pose" "noBreak"
        movej(pose_trans(easyPickPose,p[0.0000,0.0000,0.0300,0.0000,0.0000,0.0000]),a=1.3963,v=1.0472,t=0.000000,r=0.000000)
        # end: URCap Program Node
        # begin: URCap Program Node
        #   Source: SensoPart VISOR Robotic, 2.0.0, SensoPart Industriesensorik GmbH
        #   Type: Target Pose
        $ 2194 "Target Pose" "noBreak"
        movel(pose_trans(easyPickPose,p[0.0000,0.0000,-0.0000,0.0000,0.0000,0.0000]),a=0.5000,v=0.2500,t=0.000000,r=0.000000)
        # end: URCap Program Node
        $ 2195 "Close Gripper" "noBreak"
        # begin: URCap Program Node
        #   Source: Robotiq_Grippers, 1.8.4.4844, Robotiq Inc.
        #   Type: Gripper
        $ 2196 "Gripper Open (1)" "noBreak"
        if not(gripper_connected[0]):
          popup("Gripper 1 must be connected to run this program.", "No connection", False, True, True)
        end
        if not(rq_is_gripper_activated("1")):
          popup("Gripper 1 is not activated. Go to Installation tab > Gripper to activate it and run the program again.", "Not activated", False, True, True)
        end
        rq_set_pos_spd_for(0, 255, 255, "1")
        rq_wait_pos_spe_for_request(0, 255, 255, "1")
        rq_go_to("1")
        rq_wait("1")
        # end: URCap Program Node
        # begin: URCap Program Node
        #   Source: SensoPart VISOR Robotic, 2.0.0, SensoPart Industriesensorik GmbH
        #   Type: Exit Pose
        $ 2197 "Exit Pose" "noBreak"
        movel(pose_trans(easyPickPose,p[0.0000,0.0000,0.0500,0.0000,0.0000,0.0000]),a=0.5000,v=0.2500,t=0.000000,r=0.000000)
        # end: URCap Program Node
        easyPickObjTaken = True
      end
      # end: URCap Program Node
      # begin: URCap Program Node
      #   Source: SensoPart VISOR Robotic, 2.0.0, SensoPart Industriesensorik GmbH
      #   Type: No Object Detected
      $ 2198 "No Object Detected" "noBreak"
      if (visor_partsFound(easyPickVisorId) < 1):
        $ 2199 "Popup: No weigh scale detected" "noBreak"
        popup("No weigh scale detected", "Message", False, False, blocking=True)
        else:
      end
      # end: URCap Program Node
    end
    easyPickCount_1 = easyPickCount_1 + 1
    visor_easyPickUpdate(easyPickVisorId, "counter", easyPickCount_1)
    visor_easyPickSetIdent("425780", easyPickVisorId)
    # end: URCap Program Node
  end
  visorFuncEasyPick_7a8a4a()
  # end: URCap Program Node
  $ 2200 "MoveJ"
  $ 2201 "Waypoint_46" "breakAfter"
  movej(get_inverse_kin(Waypoint_46_p, qnear=Waypoint_46_q), a=1.3962634015954636, v=1.0471975511965976, r=0.05)
  $ 2202 "Waypoint_32" "breakAfter"
  movej(get_inverse_kin(Waypoint_32_p, qnear=Waypoint_32_q), a=1.3962634015954636, v=1.0471975511965976, r=0.011)
  $ 2203 "MoveL"
  $ 2204 "Waypoint_33" "breakAfter"
  movel(Waypoint_33_p, a=1.2, v=0.25, r=0.05)
  $ 2205 "Waypoint_34" "breakAfter"
  movel(Waypoint_34_p, a=1.2, v=0.25, r=0.009000000000000001)
  # begin: URCap Program Node
  #   Source: Robotiq_Grippers, 1.8.4.4844, Robotiq Inc.
  #   Type: Gripper
  $ 2206 "Gripper Move10mm (1)"
  if not(gripper_connected[0]):
    popup("Gripper 1 must be connected to run this program.", "No connection", False, True, True)
  end
  if not(rq_is_gripper_activated("1")):
    popup("Gripper 1 is not activated. Go to Installation tab > Gripper to activate it and run the program again.", "Not activated", False, True, True)
  end
  rq_set_pos_spd_for(203, 64, 62, "1")
  rq_wait_pos_spe_for_request(203, 64, 62, "1")
  rq_go_to("1")
  rq_wait("1")
  # end: URCap Program Node
  $ 2207 "MoveL"
  $ 2208 "Waypoint_40" "breakAfter"
  movel(Waypoint_40_p, a=1.2, v=0.25, r=0.001)
  $ 2209 "decap_1" "breakAfter"
  movel(decap_1_p, a=1.2, v=0.25)
  # begin: URCap Program Node
  #   Source: Robotiq_Grippers, 1.8.4.4844, Robotiq Inc.
  #   Type: Gripper
  $ 2210 "Gripper Move45mm (1)"
  if not(gripper_connected[0]):
    popup("Gripper 1 must be connected to run this program.", "No connection", False, True, True)
  end
  if not(rq_is_gripper_activated("1")):
    popup("Gripper 1 is not activated. Go to Installation tab > Gripper to activate it and run the program again.", "Not activated", False, True, True)
  end
  rq_set_pos_spd_for(40, 173, 153, "1")
  rq_wait_pos_spe_for_request(40, 173, 153, "1")
  rq_go_to("1")
  rq_wait("1")
  # end: URCap Program Node
  $ 2211 "MoveL"
  $ 2212 "Waypoint_41" "breakAfter"
  movel(Waypoint_41_p, a=1.2, v=0.25)
  $ 2213 "Waypoint_42" "breakAfter"
  movel(Waypoint_42_p, a=1.2, v=0.25)
  $ 2214 "decap_2" "breakAfter"
  movel(decap_2_p, a=1.2, v=0.25)
  # begin: URCap Program Node
  #   Source: Robotiq_Grippers, 1.8.4.4844, Robotiq Inc.
  #   Type: Gripper
  $ 2215 "Gripper Move10mm (1)"
  if not(gripper_connected[0]):
    popup("Gripper 1 must be connected to run this program.", "No connection", False, True, True)
  end
  if not(rq_is_gripper_activated("1")):
    popup("Gripper 1 is not activated. Go to Installation tab > Gripper to activate it and run the program again.", "Not activated", False, True, True)
  end
  rq_set_pos_spd_for(203, 99, 79, "1")
  rq_wait_pos_spe_for_request(203, 99, 79, "1")
  rq_go_to("1")
  rq_wait("1")
  # end: URCap Program Node
  $ 2216 "MoveL"
  $ 2217 "Waypoint_44" "breakAfter"
  movel(Waypoint_44_p, a=1.2, v=0.25)
  $ 2218 "Waypoint_45" "breakAfter"
  movel(Waypoint_45_p, a=1.2, v=0.25)
  $ 2219 "decap_1" "breakAfter"
  movel(decap_1_p, a=1.2, v=0.25)
  $ 2220 "Waypoint_35" "breakAfter"
  movel(Waypoint_35_p, a=1.2, v=0.25)
  $ 2221 "Waypoint_36" "breakAfter"
  movel(Waypoint_36_p, a=1.2, v=0.25)
  $ 2222 "Waypoint_37" "breakAfter"
  movel(Waypoint_37_p, a=1.2, v=0.25, r=0.05)
  $ 2223 "Waypoint_38" "breakAfter"
  movel(Waypoint_38_p, a=1.2, v=0.25, r=0.05)
  # begin: URCap Program Node
  #   Source: Robotiq_Grippers, 1.8.4.4844, Robotiq Inc.
  #   Type: Gripper
  $ 2224 "Gripper Move38mm (1)"
  if not(gripper_connected[0]):
    popup("Gripper 1 must be connected to run this program.", "No connection", False, True, True)
  end
  if not(rq_is_gripper_activated("1")):
    popup("Gripper 1 is not activated. Go to Installation tab > Gripper to activate it and run the program again.", "Not activated", False, True, True)
  end
  rq_set_pos_spd_for(73, 173, 153, "1")
  rq_wait_pos_spe_for_request(73, 173, 153, "1")
  rq_go_to("1")
  rq_wait("1")
  # end: URCap Program Node
  $ 2225 "MoveL"
  $ 2226 "Waypoint_37" "breakAfter"
  movel(Waypoint_37_p, a=1.2, v=0.25, r=0.05)
  $ 2227 "Home (Safe)"
  movej([-1.2302089344500047, -1.2969853503591224, -1.875639182904262, -1.539621866126728, 1.5731943360401213, -2.80099559440227], a=1.3962634015954636, v=1.0471975511965976)
  elif (37 == switch_1):
    $ 2228 "Case 37"
    $ 2229 "Detect spatula and powder transfer"
    # begin: URCap Program Node
    #   Source: SensoPart VISOR Robotic, 2.0.0, SensoPart Industriesensorik GmbH
    #   Type: VISOR Robotic App
    $ 2230 "VISOR Easy Pick"
    def visorFuncEasyPick_ff889b():
      # begin: URCap Program Node
      #   Source: SensoPart VISOR Robotic, 2.0.0, SensoPart Industriesensorik GmbH
      #   Type: Easy Pick Setup
      $ 2231 "# 1 Setup" "noBreak"
      local easyPickVisorId = 1
      local easyPickArmMounted = True
      local easyPickSetJob = True
      local easyPickJobName = "Spatula"
      local easyPickAtImgAcq = False
      local easyPickImgAcqPose = p[-0.1334,-0.4212,0.2049,-0.9203,1.0979,-1.4781]
      # end: URCap Program Node
      # begin: URCap Program Node
      #   Source: SensoPart VISOR Robotic, 2.0.0, SensoPart Industriesensorik GmbH
      #   Type: Process
      $ 2232 "Process" "noBreak"
      local easyPickObjTaken = False
      local easyPickTrigger = False
      local easyPickPoseIdx = 0
      local easyPickPose = p[0,0,0,0,0,0]
      def easyPickFuncTrigger(visorId, setJob, jobName, arm):
      if (setJob):
        visor_changeJob(visorId, jobName, 6000)
      end
      if (arm):
        visor_trigger(visorId, 6000, "arm")
      else:
        visor_trigger(visorId, 6000)
      end
      global easyPickParts_3=visor_partsFound(visorId)
      visor_easyPickUpdate(visorId, "parts", visor_partsFound(visorId))
      return visor_getPose3d(visorId, 0)
    end
    while (not easyPickObjTaken):
      easyPickTrigger = (easyPickCount_3 >= visor_partsFound(easyPickVisorId)) or (easyPickCount_3 > 9) or (not visor_easyPickCheckIdent("edc17a", easyPickVisorId))
      if (easyPickTrigger):
        easyPickCount_3 = 0
      end
      easyPickPoseIdx = easyPickCount_3
      easyPickPose = visor_getPose3d(easyPickVisorId, easyPickPoseIdx)
      visor_easyPickUpdate(easyPickVisorId, "counter", easyPickPoseIdx)
      # begin: URCap Program Node
      #   Source: SensoPart VISOR Robotic, 2.0.0, SensoPart Industriesensorik GmbH
      #   Type: Image Acquisition Pose
      $ 2233 "Image Acquisition Pose" "noBreak"
      if (easyPickTrigger):
        if (not easyPickAtImgAcq):
          movej(pose_trans(easyPickImgAcqPose,p[0.0000,0.0000,-0.0000,0.0000,0.0000,0.0000]),a=1.3963,v=1.0472,t=0.000000,r=0.000000)
          easyPickAtImgAcq = True
        end
        easyPickPose = easyPickFuncTrigger(easyPickVisorId, easyPickSetJob, easyPickJobName, easyPickArmMounted)
      end
      # end: URCap Program Node
      # begin: URCap Program Node
      #   Source: SensoPart VISOR Robotic, 2.0.0, SensoPart Industriesensorik GmbH
      #   Type: Object Detected
      $ 2234 "Object Detected" "noBreak"
      if (visor_partsFound(easyPickVisorId) > 0):
        $ 2235 "Open Gripper" "noBreak"
        # begin: URCap Program Node
        #   Source: Robotiq_Grippers, 1.8.4.4844, Robotiq Inc.
        #   Type: Gripper
        $ 2236 "Gripper Open (1)" "noBreak"
        if not(gripper_connected[0]):
          popup("Gripper 1 must be connected to run this program.", "No connection", False, True, True)
        end
        if not(rq_is_gripper_activated("1")):
          popup("Gripper 1 is not activated. Go to Installation tab > Gripper to activate it and run the program again.", "Not activated", False, True, True)
        end
        rq_set_pos_spd_for(0, 130, 89, "1")
        rq_wait_pos_spe_for_request(0, 130, 89, "1")
        rq_go_to("1")
        rq_wait("1")
        # end: URCap Program Node
        # begin: URCap Program Node
        #   Source: SensoPart VISOR Robotic, 2.0.0, SensoPart Industriesensorik GmbH
        #   Type: Approach Pose
        $ 2237 "Approach Pose" "noBreak"
        movej(pose_trans(easyPickPose,p[0.0000,0.0000,0.1000,0.0000,0.0000,0.0000]),a=1.3963,v=1.0472,t=0.000000,r=0.000000)
        # end: URCap Program Node
        # begin: URCap Program Node
        #   Source: SensoPart VISOR Robotic, 2.0.0, SensoPart Industriesensorik GmbH
        #   Type: Target Pose
        $ 2238 "Target Pose" "noBreak"
        movel(pose_trans(easyPickPose,p[0.0000,0.0000,-0.0000,0.0000,0.0000,0.0000]),a=0.5000,v=0.2500,t=0.000000,r=0.000000)
        # end: URCap Program Node
        $ 2239 "Close Gripper" "noBreak"
        # begin: URCap Program Node
        #   Source: Robotiq_Grippers, 1.8.4.4844, Robotiq Inc.
        #   Type: Gripper
        $ 2240 "Gripper Close (1)" "noBreak"
        if not(gripper_connected[0]):
          popup("Gripper 1 must be connected to run this program.", "No connection", False, True, True)
        end
        if not(rq_is_gripper_activated("1")):
          popup("Gripper 1 is not activated. Go to Installation tab > Gripper to activate it and run the program again.", "Not activated", False, True, True)
        end
        rq_set_pos_spd_for(255, 130, 89, "1")
        rq_wait_pos_spe_for_request(255, 130, 89, "1")
        rq_go_to("1")
        rq_wait("1")
        # end: URCap Program Node
        # begin: URCap Program Node
        #   Source: SensoPart VISOR Robotic, 2.0.0, SensoPart Industriesensorik GmbH
        #   Type: Exit Pose
        $ 2241 "Exit Pose" "noBreak"
        movel(pose_trans(easyPickPose,p[0.0000,0.0000,0.2000,0.0000,0.0000,0.0000]),a=0.5000,v=0.2500,t=0.000000,r=0.000000)
        # end: URCap Program Node
        easyPickObjTaken = True
      end
      # end: URCap Program Node
      # begin: URCap Program Node
      #   Source: SensoPart VISOR Robotic, 2.0.0, SensoPart Industriesensorik GmbH
      #   Type: No Object Detected
      $ 2242 "No Object Detected" "noBreak"
      if (visor_partsFound(easyPickVisorId) < 1):
        $ 2243 "Popup: No spatula is detected" "noBreak"
        popup("No spatula is detected", "Message", False, False, blocking=True)
        else:
      end
      # end: URCap Program Node
    end
    easyPickCount_3 = easyPickCount_3 + 1
    visor_easyPickUpdate(easyPickVisorId, "counter", easyPickCount_3)
    visor_easyPickSetIdent("edc17a", easyPickVisorId)
    # end: URCap Program Node
  end
  visorFuncEasyPick_ff889b()
  # end: URCap Program Node
  $ 2244 "MoveL"
  $ 2245 "Waypoint_52" "breakAfter"
  movel(Waypoint_52_p, a=1.2, v=0.25)
  $ 2246 "Waypoint_53" "breakAfter"
  movel(Waypoint_53_p, a=0.3, v=0.05)
  $ 2247 "Loop 2 times"
  Loop_2 = 0
  while (Loop_2 < 2):
    $ 2248 "Waypoint_54" "breakAfter"
    global move_thread_flag_2248=0
    thread move_thread_2248():
      enter_critical
      move_thread_flag_2248 = 1
      movel(Waypoint_54_p, a=0.3, v=0.05)
      move_thread_flag_2248 = 2
      exit_critical
    end
    move_thread_flag_2248 = 0
    move_thread_han_2248 = run move_thread_2248()
    while (True):
      local targetTcpDirection=get_target_tcp_speed()
      local stepsToRetract=tool_contact(direction=targetTcpDirection)
      if (stepsToRetract > 0):
        kill move_thread_han_2248
        stopl(3.0)
        local backTrackMovement=get_actual_joint_positions_history(stepsToRetract)
        local contactPose=get_forward_kin(backTrackMovement)
        local posDir=[targetTcpDirection[0],targetTcpDirection[1],targetTcpDirection[2]]
        local retractTo=contactPose
        if (norm(posDir) > 1e-6):
          local normalizedPosDir=normalize(posDir)
          local additionalRetraction=p[normalizedPosDir[0] * 0.0, normalizedPosDir[1] * 0.0, normalizedPosDir[2] * 0.0, 0, 0, 0]
          retractTo = pose_sub(contactPose, additionalRetraction)
        end
        movel(retractTo, a=3.0, v=0.1)
        $ 2249 "Until (tool_contact_detection)"
        break
      end
      sleep(1.0E-10)
      if (move_thread_flag_2248 > 1):
        join move_thread_han_2248
        break
      end
      sync()
    end
    $ 2250 "Waypoint_55" "breakAfter"
    movel(Waypoint_55_p, a=0.3, v=0.05)
    $ 2251 "Waypoint_56" "breakAfter"
    movel(Waypoint_56_p, a=0.3, v=0.05)
    Loop_2 = Loop_2 + 1
  end
  $ 2252 "Waypoint_57" "breakAfter"
  movel(Waypoint_57_p, a=1.5, v=0.75)
  $ 2253 "Waypoint_56" "breakAfter"
  movel(Waypoint_56_p, a=0.3, v=0.05, r=0.016999999999999998)
  $ 2254 "Waypoint_58" "breakAfter"
  movel(Waypoint_58_p, a=0.3, v=0.05, r=0.05)
  $ 2255 "Waypoint_59" "breakAfter"
  movel(Waypoint_59_p, a=0.3, v=0.05, r=0.05)
  $ 2256 "Waypoint_60" "breakAfter"
  movel(Waypoint_60_p, a=1.2, v=0.25, r=0.05)
  $ 2257 "Waypoint_61" "breakAfter"
  movel(Waypoint_61_p, a=1.2, v=0.25, r=0.05)
  $ 2258 "Waypoint_62" "breakAfter"
  movel(Waypoint_62_p, a=1.2, v=0.25)
  $ 2259 "Waypoint_63" "breakAfter"
  global move_thread_flag_2259=0
  thread move_thread_2259():
    enter_critical
    move_thread_flag_2259 = 1
    movel(Waypoint_63_p, a=0.1, v=0.02)
    move_thread_flag_2259 = 2
    exit_critical
  end
  move_thread_flag_2259 = 0
  move_thread_han_2259 = run move_thread_2259()
  while (True):
    sleep(1.0E-10)
    if (move_thread_flag_2259 > 1):
      join move_thread_han_2259
      break
    end
    sync()
  end
  end
  $ 2278 "'=========='"
  # '=========='
  $ 2279 "PostSettings"
  $ 2280 "'ADD ADDITIONAL CHECKS'"
  # 'ADD ADDITIONAL CHECKS'
  end
  $ 2 "BeforeStart"
  $ 3 "Scripts"
  $ 4 "Script: 001 SCRIPT Errors and Warnings Deifnes V0.2.script"

  #*****************************************************
  # customer          :   UK Essen
  # project name      :   P1132
  #****************************************************
  # controller        :
  # software          :
  #****************************************************
  # author            :   E.Petrichenko
  # Copyright (c)     :   United Robotics Group Health and Food GmbH
  #                       An der Riede 2
  #                       28816 Stuhr
  #                       Germany
  #****************************************************
  # description       :   centrifuge actions for the application
  # version:      	:   0.1
  # created           :   22.08.2024
  # updated           :
  #****************************************************
  # modifications     :
  #
  # date              :
  # name              :
  # reason            :
  #****************************************************


  #################################### VARIABLES DEFINITIONS ###################################

  ERROR_POSE_NOT_REACHABLE = 1002
  ERROR_ROBOT_ARM_NOT_IN_HOME_POSE = 1006
  ERROR_NO_OBJECT_TO_PICK = 1010
  ERROR_NOT_DOCKED = 2003
  ERROR_NOT_REACHABLE_TARGET = 2007
  ERROR_CHARGING_NOT_STARTED = 2008
  ERROR_AMR_WRONG_MODE = 2009
  ERROR_UNKNOWN_POSE = 2010
  ERROR_NO_LANDMARK = 3002
  ERROR_WRONG_ORDER = 4002
  ERROR_CENTRIFUGE_CONNECTION = 5001
  ERROR_CENTRIFUGE_POWER = 5002
  ERROR_CENTRIFUGE = 5003
  ERROR_CENTRIFUGE_LID = 5004
  ERROR_CANNOT_OPEN_HATCH = 5006
  ERROR_CANNOT_CLOSE_HATCH = 5008
  ERROR_CANNOT_ROTATE = 5010
  ERROR_CANNOT_START = 5011
  ERROR_WRONG_KEY_POSE = 5012
  ERROR_MISSIING_CENTRACK = 5013

  WARNING_POSE_NOT_REACHABLE = 1002
  WARNING_BATTERY_LEVEL = 2002
  WARNING_NOT_REACHABLE_TARGET = 2007


  ERROR = struct(
      FLAG = False,
      ID = 0,
      MSG = "")

  WARNING = struct(
      FLAG = False,
      ID = 0,
      MSG = "")


  #################################### FUNCTIONS ###################################

  def set_error(error_id):
      ERROR.ID = error_id
      if (ERROR.ID == 0):
          ERROR.FLAG = False
          ERROR.MSG = ""
      else:
          ERROR.FLAG = True
          if(ERROR.ID == ERROR_POSE_NOT_REACHABLE):
              ERROR.MSG = "Pose is not reachable"
          elif(ERROR.ID == ERROR_NO_OBJECT_TO_PICK):
              ERROR.MSG = "No object to pick"
          elif(ERROR.ID == ERROR_NO_LANDMARK):
              ERROR.MSG = "No landmark detected"
          elif(ERROR.ID == ERROR_ROBOT_ARM_NOT_IN_HOME_POSE):
              ERROR.MSG = "Robot arm cannot go to home pose"
          elif(ERROR.ID == ERROR_AMR_WRONG_MODE):
              ERROR.MSG = "AMR is in the wrong mode"
          elif(ERROR.ID == ERROR_NOT_DOCKED):
              ERROR.MSG = "Could not dock to the charger"
          elif(ERROR.ID == ERROR_NOT_REACHABLE_TARGET):
              ERROR.MSG = "Could not reach the target"
          elif(ERROR.ID == ERROR_CHARGING_NOT_STARTED):
              ERROR.MSG = "Could not start charging"
          elif(ERROR.ID == ERROR_UNKNOWN_POSE):
              ERROR.MSG = "Unknown navigation target"
          elif(ERROR.ID == ERROR_CANNOT_OPEN_HATCH):
              ERROR.MSG = "Centrifuge Cannot open the hatch"
          elif(ERROR.ID == ERROR_CENTRIFUGE_CONNECTION):
              ERROR.MSG = "Cannot reach centrifuge"
          elif (ERROR.ID == ERROR_CANNOT_CLOSE_HATCH):
              ERROR.MSG = "Centrifuge Cannot close the hatch"
          elif (ERROR.ID == ERROR_CANNOT_START):
              ERROR.MSG = "Centrifuge Cannot start"
          elif (ERROR.ID == ERROR_CANNOT_ROTATE):
              ERROR.MSG = "Centrifuge Cannot rotate the rotor"
          elif (ERROR.ID == ERROR_WRONG_ORDER):
              ERROR.MSG = "Wrong parameter was recieved"
          elif (ERROR.ID == ERROR_CENTRIFUGE):
              ERROR.MSG = "Centrifuge is in Error"
          elif (ERROR.ID == ERROR_WRONG_KEY_POSE):
              ERROR.MSG = "Key is in the wrong position"
          elif(ERROR.ID == ERROR_MISSIING_CENTRACK):
              ERROR.MSG = "Missing rack for centrifuge set"
          elif(ERROR.ID == ERROR_CENTRIFUGE_POWER):
              ERROR.MSG = "Centrifuge is turned off"
          elif(ERROR.ID == ERROR_CENTRIFUGE_LID):
              ERROR.MSG = "Lid of the centrifuge is opened"
          else:
              ERROR.MSG = "Unknown code"
          end
          textmsg("ERROR:",ERROR)
      end
  end

  def set_warning(warning_id):
      WARNING.ID = warning_id
      if (WARNING.ID == 0):
          WARNING.FLAG = False
          WARNING.MSG = ""
      else:
          WARNING.FLAG = True
          if(WARNING.ID == WARNING_POSE_NOT_REACHABLE):
              WARNING.MSG = "Pose is not reachable"
          elif(WARNING.ID == WARNING_BATTERY_LEVEL):
              WARNING.MSG = "Batery level dropped to a certain level"
          elif(WARNING.ID == WARNING_NOT_REACHABLE_TARGET):
              WARNING.MSG = "Not reachable location of AMR"
          else:
              WARNING.MSG = "Unknown code"
          end
          textmsg("WARNING:",WARNING)
      end
  end


  def reset_error():
    ERROR.ID = 0
    ERROR.FLAG = False
    ERROR.MSG = ""
  end


  def reset_warning():
      WARNING.ID = 0
      WARNING.FLAG = False
      WARNING.MSG = ""
    end
  $ 5 "Script: SCRIPT uGO V7.11.1.script"
  #*****************************************************
  # customer          :
  # project name      :   Standard Application
  #****************************************************
  # controller        :
  # software          :
  #****************************************************
  # author            :   P. Koehnke
  # Copyright (c)     :   United Robotics Group
  #                       An der Riede 2
  #                       28816 Stuhr
  #                       Germany
  #****************************************************
  # description       :   interface for uGo
  # version:      	:   6.0
  # created           :   21.04.2022
  # updated           :
  #****************************************************
  # modifications     :   add new rpc-functions to interchange more data
  #
  # date              :   2024-02-29
  # name              :   P. Koehnke
  # reason            :   implemtentation of PackML behavoiur in uGO
  #****************************************************
  #****************************************************
  # modifications     :   add reflecting the UID of the uGO task back to uGO
  #
  # date              :   2024-07-02
  # name              :   P. Koehnke
  # reason            :   be sure to finish the right tasks
  #****************************************************

  # available rpc-functions:
  #.on('con_check', (err, _params, callback) => callback(err, this.con_check()))
  #.on('read_input', (err, params, callback) => callback(err, this.read_input(params[0], params[1])))
  #.on('write_output', (err, params, callback) => callback(err, this.write_output(params[0], params[1], params[2])))
  #.on('read_status', (err, params, callback) => callback(err, this.read_status(params[0])))
  #.on('write_status', (err, params, callback) => callback(err, this.write_status(params[0], params[1])))
  #.on('send_template', (err, params, callback) => callback(err, this.receive_state(params[0])))
  #.on('receive_event', (err, params, callback) => callback(err, this.send_event()))
  #.on('send_state', (err, params, callback) => callback(err, this.receive_state(params[0])))
  #.on('send_error', (err, params, callback) => callback(err, this.receive_error(params[0])))
  #.on('NotFound', (methodCalled, params) => LOG.warn('Method "', methodCalled, '" does not exist. ', { params }));

  # =======================================================================
  local IDX_CMD_STOP = 0
  local IDX_CMD_RESET = 1
  local IDX_CMD_START = 2
  local IDX_CMD_HOLD = 3
  local IDX_CMD_UNHOLD = 4
  local IDX_CMD_SUSPEND = 5
  local IDX_CMD_UNSUSPEND = 6
  local IDX_CMD_ABORT = 7
  local IDX_CMD_CLEAR = 8
  local IDX_FNC_FREEDRIVE = 9

  # uGo specific declarations
  global UGO_Request_ID = ""
  global UGO_UNIT_Task = ""
  global UGO_Task_ID = 0
  global UGO_Event = ""
  local UGO_Enable_Control = False
  local UGO = rpc_factory("xmlrpc", "http://192.168.12.120:8080")
  local UGO_Ctrl_Cmd = [False, False, False, False, False, False, False, False, False, False]

  local UGO_AMR_Pos = struct(position_identifier=0, x1=0, x2=0, y1=0, y2=0, theta1=0, theta2=0)
  local UGO_EOAT = struct(object_picked=False)

  def ugo_init(enable=True, rpc_address="http://192.168.12.120:8080"):
      # connection with uGo
      if enable:
          UGO = rpc_factory("xmlrpc", rpc_address)
          UGO_Enable_Control = True
      else:
          UGO_Enable_Control = False
      end
  end

  def ugo_event_controller():
      # interpret the given command and map it to the internal commands
      if UGO_Enable_Control:
          UGO_Event = UGO.receive_event()
      end

      UGO_Ctrl_Cmd[IDX_CMD_STOP] = (UGO_Event == "stop")
      UGO_Ctrl_Cmd[IDX_CMD_RESET] = (UGO_Event == "reset")
      UGO_Ctrl_Cmd[IDX_CMD_START] = (UGO_Event == "start")
      UGO_Ctrl_Cmd[IDX_CMD_HOLD] = (UGO_Event == "hold")
      UGO_Ctrl_Cmd[IDX_CMD_UNHOLD] = (UGO_Event == "un_hold")
      UGO_Ctrl_Cmd[IDX_CMD_SUSPEND] = (UGO_Event == "suspend")
      UGO_Ctrl_Cmd[IDX_CMD_UNSUSPEND] = (UGO_Event == "un_suspend")
      UGO_Ctrl_Cmd[IDX_CMD_ABORT] = (UGO_Event == "abort")
      UGO_Ctrl_Cmd[IDX_CMD_CLEAR] = (UGO_Event == "clear")
      UGO_Ctrl_Cmd[IDX_FNC_FREEDRIVE] = (UGO_Event == "freedrive")

      return UGO_Ctrl_Cmd
  end

  def ugo_translate_pml_state():
      # translate the current PML State to a string
      if (STATE == 1):
          return "STOPPING"
      elif (STATE == 2):
          return "STOPPED"
      elif (STATE == 3):
          return "RESETTING"
      elif (STATE == 4):
          return "IDLE"
      elif (STATE == 5):
          return "STARTING"
      elif (STATE == 6):
          return "EXECUTE"
      elif (STATE == 7):
          return "COMPLETING"
      elif (STATE == 8):
          return "COMPLETE"
      elif (STATE == 9):
          return "HOLDING"
      elif (STATE == 10):
          return "HELD"
      elif (STATE == 11):
          return "UNHOLDING"
      elif (STATE == 12):
          return "SUSPENDING"
      elif (STATE == 13):
          return "SUSPENDED"
      elif (STATE == 14):
          return "UNSUSPENDING"
      elif (STATE == 15):
          return "ABORTING"
      elif (STATE == 16):
          return "ABORTED"
      elif (STATE == 17):
          return "CLEARING"
      else:
          return "UNKNOWN"
      end
  end

  def ugo_update_outputs():
      #Update the outputs to uGo via xmplrpc service
      UGO.write_status("ROB_Skill", UGO_UNIT_Task)
      UGO.write_status("ROB_Battery", AMR_Battery)
      UGO.write_status("ROB_Gripper", OBJ_Picked)
      UGO.send_state(ugo_translate_pml_state(), UGO_UNIT_Task)
      UGO.send_error(ERROR.ID)
      #UGO.send_position(AMR_Position)
  end

  def ugo_get_task():
      # get the actual task to work on
      # added: reflecting the UID of the task back to uGO
      UGO_UNIT_Task = UGO.read_status("DSH_Workflow")
      if (UGO_UNIT_Task != ""):
          UGO_Request_ID = str_sub(UGO_UNIT_Task, 0, 39)
          UGO_Task_ID = to_num(str_sub(UGO_UNIT_Task, 40, 2))
          #ugo_tasks()
          return UGO_Task_ID
      else:
          return 0
      end
  end

  def ugo_pml_stopping():
      return True
  end

  def ugo_pml_resetting():
      ugo_get_task()
      if (UGO_UNIT_Task == ""):
          UGO_Request_ID = ""
          UGO_Task_ID = 0
          return True
      end
      return False
  end

  def ugo_pml_starting():
      #UGO_Task_Content = UGO.receive_task()
      return (UGO_UNIT_Task != "")
  end

  def ugo_pml_holding():
      return True
  end

  def ugo_pml_unholding():
      return True
  end

  def ugo_pml_suspending():
      return True
  end

  def ugo_pml_unsuspending():
      return True
  end

  def ugo_pml_completing():
      return True
  end

  def ugo_pml_aborting():
      return True
  end

  def ugo_pml_clearing():
      return True
  end

  # =======================================================================
  # end of uGO script
  # =======================================================================
  $ 7 "Script: SCRIPT PackML V1.2.1.script"
  # PackML

  IO_ADDRESS_CMD_STOP = 1
  IO_ADDRESS_CMD_RESET = 7
  IO_ADDRESS_CMD_START = 0

  EXT_ADDRESS_CMD_STOP = 0
  EXT_ADDRESS_CMD_RESET = 1
  EXT_ADDRESS_CMD_START = 2
  EXT_ADDRESS_CMD_HOLD = 3
  EXT_ADDRESS_CMD_UNHOLD = 4
  EXT_ADDRESS_CMD_SUSPEND = 5
  EXT_ADDRESS_CMD_UNSUSPEND = 6
  EXT_ADDRESS_CMD_ABORT = 7
  EXT_ADDRESS_CMD_CLEAR = 8
  EXT_ADDRESS_FNC_FREEDRIVE = 9

  global EXT_CtrlCmd = [False, False, False, False, False, False, False, False, False, False]

  EXT_Control_by = "uGO"

  global CMD_Abort = False
  global CMD_Clear = False
  global CMD_Stop = False
  global CMD_Reset = False
  global CMD_Start = False
  global CMD_Hold = False
  global CMD_Unhold = False
  global CMD_Suspend = False
  global CMD_Unsuspend = False
  global FNC_Freedrive = False

  CND_Suspend = False         # condition for suspend command
  CND_Unsuspend = False       # condition for unsuspend command

  thread Get_Pml_Command():
      while (True):
          if (EXT_Control_by == "uGO"):
              EXT_CtrlCmd = ugo_event_controller()
          elif (EXT_Control_by == "Leitsystem"):
              # EXT_CtrlCmd = Leitsystem
          end
          # ---------- Abort ---------- #
          if ((not STATE == 15) and (not STATE == 16) and EXT_CtrlCmd[EXT_ADDRESS_CMD_ABORT]):
              CMD_Abort = True
              CMD_Stop = False
          elif ((STATE == 17) and not EXT_CtrlCmd[EXT_ADDRESS_CMD_ABORT]):
              CMD_Abort = False
          end
          # ---------- Stop ---------- #
          if ((not STATE == 1) and (not STATE == 2) and (get_standard_digital_in(IO_ADDRESS_CMD_STOP) or EXT_CtrlCmd[EXT_ADDRESS_CMD_STOP])):
              CMD_Stop = True
              if get_standard_digital_in(IO_ADDRESS_CMD_STOP):
                  log_state("Stop command by pushbutton")
              elif EXT_CtrlCmd[EXT_ADDRESS_CMD_STOP]:
                  log_state("Stop command by external control")
              end
          elif (STATE == 2) and (not get_standard_digital_in(IO_ADDRESS_CMD_STOP)) and (not EXT_CtrlCmd[EXT_ADDRESS_CMD_STOP]):
              CMD_Stop = False
          end
          CMD_Hold = (STATE == 6 or STATE == 10) and not CMD_Stop and (ERROR.FLAG or EXT_CtrlCmd[EXT_ADDRESS_CMD_HOLD])
          CMD_Reset = (STATE == 2 or STATE == 8) and not CMD_Stop and (read_input_boolean_register(5) or EXT_CtrlCmd[EXT_ADDRESS_CMD_RESET])
          CMD_Start = (STATE == 4) and not CMD_Stop and (get_standard_digital_in(IO_ADDRESS_CMD_START) or EXT_CtrlCmd[EXT_ADDRESS_CMD_START])
          CMD_Unhold = (STATE == 10) and not CMD_Stop and (get_standard_digital_in(IO_ADDRESS_CMD_START) or EXT_CtrlCmd[EXT_ADDRESS_CMD_UNHOLD])
          CMD_Suspend = (STATE == 6) and not CMD_Stop and (CND_Suspend or EXT_CtrlCmd[EXT_ADDRESS_CMD_SUSPEND])
          CMD_Unsuspend = (STATE == 13) and not CMD_Stop and (CND_Unsuspend or EXT_CtrlCmd[EXT_ADDRESS_CMD_UNSUSPEND])
          CMD_Clear = (STATE == 16) and EXT_CtrlCmd[EXT_ADDRESS_CMD_CLEAR]
          FNC_Freedrive = (STATE == 10) and EXT_CtrlCmd[EXT_ADDRESS_FNC_FREEDRIVE]
          sleep(0.1)
      end
  end

  thread_pml_command_handler = run Get_Pml_Command()

  def command_manager(external_control="uGO", cond_suspend=False, cond_unsuspend=False):

      EXT_Control_by = external_control
      CND_Suspend = cond_suspend
      CND_Unsuspend = cond_unsuspend

      if (CMD_Abort and STATE != 15 and STATE != 16):
          STATE = 15
      elif (CMD_Stop and STATE != 1 and STATE != 2):
          STATE = 1
      end
      return False
  end

  def stopping():
      if (EXT_Control_by == "uGO"):
          return ugo_pml_stopping()
      elif (EXT_Control_by == "Leitsystem"):
          # EXT_CtrlCmd = Leitsystem
      else:
          return True
      end
      return False
  end

  def resetting():
      if (EXT_Control_by == "uGO"):
          return ugo_pml_resetting()
      elif (EXT_Control_by == "Leitsystem"):
          # EXT_CtrlCmd = Leitsystem
      else:
          return True
      end
      return False
  end

  def starting():
      if (EXT_Control_by == "uGO"):
          return ugo_pml_starting()
      elif (EXT_Control_by == "Leitsystem"):
          # EXT_CtrlCmd = Leitsystem
      else:
          return True
      end
      return False
  end

  def holding():
      if (EXT_Control_by == "uGO"):
          return ugo_pml_holding()
      elif (EXT_Control_by == "Leitsystem"):
          # EXT_CtrlCmd = Leitsystem
      else:
          return True
      end
      return False
  end

  def unholding():
      if (EXT_Control_by == "uGO"):
          return ugo_pml_unholding()
      elif (EXT_Control_by == "Leitsystem"):
          # EXT_CtrlCmd = Leitsystem
      else:
          return True
      end
      return False
  end

  def suspending():
      if (EXT_Control_by == "uGO"):
          return ugo_pml_suspending()
      elif (EXT_Control_by == "Leitsystem"):
          # EXT_CtrlCmd = Leitsystem
      else:
          return True
      end
      return False
  end

  def unsuspending():
      if (EXT_Control_by == "uGO"):
          return ugo_pml_unsuspending()
      elif (EXT_Control_by == "Leitsystem"):
          # EXT_CtrlCmd = Leitsystem
      else:
          return True
      end
      return False
  end

  def completing():
      if (EXT_Control_by == "uGO"):
          return ugo_pml_completing()
      elif (EXT_Control_by == "Leitsystem"):
          # EXT_CtrlCmd = Leitsystem
      else:
          return True
      end
      return False
  end

  def aborting():
      if (EXT_Control_by == "uGO"):
          return ugo_pml_aborting()
      elif (EXT_Control_by == "Leitsystem"):
          # EXT_CtrlCmd = Leitsystem
      else:
          return True
      end
      return False
  end

  def clearing():
      if (EXT_Control_by == "uGO"):
          return ugo_pml_clearing()
      elif (EXT_Control_by == "Leitsystem"):
          # EXT_CtrlCmd = Leitsystem
      else:
          return True
      end
      return False
  end
  $ 8 "Script: SCRIPT Utility V5.5.script"
  #*****************************************************
  # customer          :   tbd
  # project name      :   tbd
  #****************************************************
  # controller        :
  # software          :
  #****************************************************
  # author            :   P. Koehnke (+49 1628859904; p.koehnke@unitedrobotics.group)
  # Copyright (c)     :   United Robotics Group Health and Food GmbH
  #                       An der Riede 2
  #                       28816 Stuhr
  #                       Germany
  #****************************************************
  # description       :   utility programs for the application
  # version:      	:   3.1
  # created           :   30.01.2023
  # updated           :
  #****************************************************
  # modifications     :   get_tool_free_pose_2(), get_index_from_list()
  #
  # date              :   05.01.2024
  # name              :   PK
  # reason            :
  #****************************************************

  def found_in_matrix(data, req_id, req_idx):
      local id = -1
      local dimensions = size(data)
      local loop_dataset = 0

      while (id != req_id and loop_dataset < dimensions[0]):
          id = data[loop_dataset, 0]
          if (id == req_id):
              return data[loop_dataset, req_idx]
          else:
              loop_dataset = loop_dataset + 1
          end
      end
  end

  def found_in_list(value, list):
      local idx = 0

      while (idx < length(list)):
          if (value == list[idx]):
              return True
          end
          idx = idx + 1
      end
      return False
  end

  def get_index_from_list(list, value = -1):
      local idx = 0

      while (idx < length(list)):
          if (value == -1):
              if (list[idx] != 0):
                  return idx
              end
          else:
              if (list[idx] == value):
                  return idx
              end
          end
          idx = idx + 1
      end
      return -1
  end

  def find_object_by_type(list, type=0):
      local object = list[0]
      local i = 0

      while i < length(list):
          object = list[i]
          if object.type == type:
              return object
          end
          i = i + 1
      end
  end

  def pose_RPY2RotVec(pose):
      local rotvec = rpy2rotvec([d2r(pose[3]), d2r(pose[4]), d2r(pose[5])])
      return p[pose[0], pose[1], pose[2], rotvec[0], rotvec[1], rotvec[2]]
  end

  def pose_RotVec2RPY(pose):
      local rpy = rotvec2rpy([pose[3], pose[4], pose[5]])
      return p[pose[0], pose[1], pose[2], r2d(rpy[0]), r2d(rpy[1]), r2d(rpy[2])]
  end

  def swivel(frame_ref, angles = [0, 0, 0], pose = p[0, 0, 0, 0, 0, 0]):

      local rpy_ref = [0, 0, 0]
      local rpy_new = [0, 0, 0]
      local rotvec_new = [0, 0, 0]
      local pose_from = p[0, 0, 0, 0, 0, 0]
      local pose_to = p[0, 0, 0, 0, 0, 0]
      local i = 0

      if (pose == p[0, 0, 0, 0, 0, 0]):
          pose_to = pose_trans(pose_inv(frame_ref), get_actual_tcp_pose())
      else:
          pose_to = pose
      end

      rpy_ref = rotvec2rpy(frame_ref[3], frame_ref[4], frame_ref[5])

      while (i < 3):
          rpy_new[i] = rpy_ref[i] + d2r(angles[i])
          i = i + 1
      end

      rotvec_new = rpy2rotvec(rpy_new)
      pose_from = p[0, 0, 0, rotvec_new[0], rotvec_new[1], rotvec_new[2]]
      pose_to = p[pose_to[0], pose_to[1], pose_to[2], rotvec_new[0], rotvec_new[1], rotvec_new[2]]

      return pose_trans(pose_from, pose_to)
  end

  def get_random_pose(pose_ref, mode = "", range_max = [0, 0, 0]):
      # modi: "cubic", "rotation"
      # getting a random pose in the x/y-plane. range can be set for each
      # translation and rotation.
      local rpy_random = [0, 0, 0]
      local rotvec_random = [0, 0, 0]
      local pose_random = pose_ref
      local i = 0

      if (mode == "cubic"):
          # cubic mode: random pose takes only x, y and z
          i = 0
          while (i < 3):
              pose_random[i] = pose_ref[i] + range_max[i] * (random() - 0.5)
              i = i + 1
          end
          return pose_random

      elif (mode == "rotation"):
          i = 0
          while (i < 3):
              rpy_random[i] = d2r(range_max[i]) * (random() - 0.5)
              i = i + 1
          end
          rotvec_random = rpy2rotvec(rpy_random)
          pose_random = pose_trans(p[0, 0, 0, rotvec_random[0], rotvec_random[1], rotvec_random[2]], pose_ref)
          return pose_random

      else:
          # unknown mode, return pose_ref
          return pose_ref
      end
  end

  def get_pattern_pos_rectangle(counter, direction, pattern, patterninc = [0, 0], patternsize = [0, 0]):
      # defines the position inside a rectangular pattern
      # pattern describes, how many objects are in x-direction and how many in y-direction [x, y]
      # patternsize will give the total length of each direction [x, y]
      local X_Fac = 0
      local Y_Fac = 0
      local max = pattern[0] * pattern[1]
      local i = 0

      if (1 > counter or counter > max):
          counter = 1
      end

      if pattern[0] == 0:
          pattern[0] = 1
      end

      if pattern[1] == 0:
          pattern[1] = 1
      end

      if (direction == "Y" or direction == "y"):
          X_Fac = floor((counter - 1) / pattern[1])
          Y_Fac = (counter - 1) % pattern[1]
      elif (direction == "X" or direction == "x"):
          X_Fac = (counter - 1) % pattern[0]
          Y_Fac = floor((counter - 1) / pattern[0])
      end

      if patternsize != [0, 0]:
          while i < 2:
              if pattern[i] > 1:
                  patterninc[i] = patternsize[i] / (pattern[i] - 1)
              end
              i = i + 1
          end
      end

      return p[X_Fac * patterninc[0], Y_Fac * patterninc[1], 0, 0, 0, 0]
  end

  def get_pattern_pos_circle(counter, radius, angle, direction, pattern, patternsize = [0, 0]):
      # get the patternpos for a circular pattern through a counter
      # need the radius and the angle in radiants
      local X_Fac = 0
      local Y_Fac = 0
      local rad_bow = 0
      local radius_cal = 0
      local ref = p[0, 0, 0, 0, 0, 0]

      if pattern[0] == 0:
          pattern[0] = 1
      end

      if pattern[1] == 0:
          pattern[1] = 1
      end

      if (direction == "Y" or direction == "y"):
          X_Fac = floor((counter - 1) / pattern[1])
          Y_Fac = (counter - 1) % pattern[1]
      elif (direction == "X" or direction == "x"):
          X_Fac = (counter - 1) % pattern[0]
          Y_Fac = floor((counter - 1) / pattern[0])
      end

      # the opening angle will be calculated in x-direction
      # works only between -90 and 90 degree
      if pattern[0] > 1:
          rad_bow = - angle / (pattern[0] - 1) * X_Fac + angle / 2
      end

      if (counter % 2 == 0 and pattern[1] > 1):
          radius_cal = radius - patternsize[1] / (pattern[1])
      else:
          radius_cal = radius + patternsize[1] / (pattern[1])
      end
      ref = p[0, radius_cal, 0, 0, 0, 0]

      return p[ref[0] * cos(rad_bow) - ref[1] * sin(rad_bow), (ref[0] * sin(rad_bow) + ref[1] * cos(rad_bow)) - radius, 0, 0, 0, 0]
  end

  def get_pattern_counter(pose, direction, pattern, patterninc = [0, 0], patternsize = [0, 0]):
      # returns the counter for a pattern from a given cartesian pose
      local patternpose = p[pose[0], pose[1], 0, 0, 0, 0]
      local X_Fac = 0
      local Y_Fac = 0
      local i = 0

      if patternsize != [0, 0]:
          while i < 2:
              if pattern[i] > 1:
                  patterninc[i] = patternsize[i] / (pattern[i] - 1)
              else:
                  pattern[i] = 0
              end
              i = i + 1
          end
      end

      # calculation of the counter in the desired axis-direction
      if (direction == "x" or direction == "X"):
          if patterninc[0] > 0:
              X_Fac = ceil((patternpose[0] + patterninc[0] / 2) / patterninc[0])
              if X_Fac < 0:
                  X_Fac = 0
              end
          end
          if patterninc[1] > 0:
              Y_Fac = floor((patternpose[1] + patterninc[1] / 2) / patterninc[1])
              if Y_Fac < 0:
                  Y_Fac = 0
            end
          end
          return Y_Fac * pattern[0] + X_Fac
      elif (direction == "y" or direction == "Y"):
          if patterninc[0] > 0:
              X_Fac = floor((patternpose[0] + patterninc[0] / 2) / patterninc[0])
          end
          if patterninc[1] > 0:
              Y_Fac = ceil((patternpose[1] + patterninc[1] / 2) / patterninc[1])
          end
          return X_Fac * pattern[1] + Y_Fac
      end
  end

  def get_plc_reg(mod_sig_name):
      return integer_to_binary_list(modbus_get_signal_status(mod_sig_name))
  end

  def set_plc_reg(mod_sig_name, mod_sig_list):
      modbus_set_output_register(mod_sig_name, binary_list_to_integer(mod_sig_list), False)
  end

  def check_decapping(offset = 0, timeout = 5, abort = False):
      # checken, ob der Deckel schon ab ist
      local start = get_actual_tcp_pose()
      local current_offset = 0
      local timecounter = 0
      while (current_offset < offset and not abort):
          current_offset = pose_dist(start, get_actual_tcp_pose())
          timecounter = timecounter + 1
          if (timecounter * 0.5 == timeout):
              break
          end
          sleep(0.5)
      end
      stopl(0.5)
  end

  def check_capping(torque = 0):
      # checken, wann der Deckel verschraubt ist
      force_mode(get_actual_tcp_pose(), [0, 0, 1, 0, 0, 0], [0, 0, -2.0, 0, 0, 0], 2, [0.01, 0.01, 0.001, 0.01, 0.01, 0.01])
  end

  def is_reachable(frame, poses, offsets = [0, 0, 0]):
      local idx = 0
      local pose = p[0, 0, 0, 0, 0, 0]

      while (idx < length(poses)):
          pose = poses[idx]
          pose[0] = pose[0] + offsets[0]
          pose[1] = pose[1] + offsets[1]
          pose[2] = pose[2] + offsets[2]

          if pose != p[0, 0, 0, 0, 0, 0]:
              if (not get_inverse_kin_has_solution(pose_trans(frame, pose))):
                  textmsg(str_cat(str_cat("Pose ", to_str(idx + 1)), " is not reachable"))
                  return False
              end
          end
          idx = idx + 1
      end
      return True
  end

  def is_within_limits(frame, poses, offsets = [0, 0, 0]):
      local idx = 0
      local pose = p[0, 0, 0, 0, 0, 0]

      while (idx < length(poses)):
          pose = poses[idx]
          pose[0] = pose[0] + offsets[0]
          pose[1] = pose[1] + offsets[1]
          pose[2] = pose[2] + offsets[2]

          if is_reachable(frame = frame, poses = poses, offsets = offsets):
              if (not is_within_safety_limits(get_inverse_kin(pose_trans(frame, pose), get_actual_joint_positions()))):
                  textmsg(str_cat(str_cat("Pose ", to_str(idx + 1)), "is out of joint limits"))
                  return False
              else:
                  idx = idx + 1
              end
          else:
              return False
          end
      end
      return True
  end


  def string_to_list(string, separator = "," , endDelimiter = ";" , capacity = 50):
      local string_length = str_len(string)
      local list_out = make_list(length = elements_in_string(string), initial_value = -1, capacity = capacity)
      local cnt = 0
      local idx = 0

      while cnt < string_length-1 :
        textmsg("new loop")
        textmsg(to_str(idx))
        local sepAt = str_find(string, separator, cnt)
        textmsg(to_str(sepAt))
        if sepAt < 0 :
            sepAt = str_find(string, endDelimiter, cnt)
        end
        list_out[idx] = to_num(str_sub(string, cnt, sepAt-cnt))
        idx = idx +1
        cnt = sepAt + 1
      end

      return list_out
  end

  def elements_in_string(string, separator = "," , endDelimiter = ";" , capacity = 50):
     local string_length = str_len(string)
      local len = 0
      local sepAt = 0

      while sepAt < string_length-1 and sepAt>=0 :
        local sepAt = str_find(string, separator, sepAt+1)
        len = len +1
      end

      return len
  end
  $ 9 "Script: SCRIPT uML Lights V1.2.script"

  #****************************************************
  # product           : uLabMobile
  # language          : urscript
  #****************************************************
  # author            :   D.Kreugel
  # Copyright (c)     :   United Robotics Group
  #                       An der Riede 2
  #                       28816 Stuhr
  #                       Germany
  #****************************************************
  # description       :   led controls for uLabMobile
  # version:      	:   1.2
  # created           :   09.08.2024
  # updated           :
  #****************************************************
  # modifications     :   changed conditions to switch lights (not only pml state but also charging state)
  #
  # date              :   09.08.2024
  # name              :   PK
  # reason            :   due to the change in project P1117, we run to often through every state. This leads to to much colorchanges
  #****************************************************

  # HARDWARE CONFIGURATION
  LED_GREEN = struct(type="CO",id=5)
  LED_RED = struct(type="CO",id=6)
  LED_BLUE = struct(type="CO",id=7)

  def set_output(type,id,state=True):
      if(type=="CO"):
          set_configurable_digital_out(id,state)
      elif(type=="DO"):
          set_standard_digital_out(id,state)
      end
  end

  def led_red_on():
      set_output(LED_RED.type,LED_RED.id,True)
  end

  def led_red_off():
      set_output(LED_RED.type,LED_RED.id,False)
  end

  def led_green_on():
      set_output(LED_GREEN.type,LED_GREEN.id,True)
  end

  def led_green_off():
      set_output(LED_GREEN.type,LED_GREEN.id,False)
  end

  def led_blue_on():
      set_output(LED_BLUE.type,LED_BLUE.id,True)
  end

  def led_blue_off():
      set_output(LED_BLUE.type,LED_BLUE.id,False)
  end


  # COLOR MIX
  def color_blue():
      led_blue_on()
      led_green_off()
      led_red_off()
  end

  def color_red():
      led_blue_off()
      led_green_off()
      led_red_on()
  end

  def color_green():
      led_blue_off()
      led_green_on()
      led_red_off()
  end

  def color_yellow():
      led_blue_off()
      led_green_on()
      led_red_on()
  end

  def color_lightblue():
      led_blue_on()
      led_green_on()
      led_red_off()
  end

  def color_violet():
      led_blue_on()
      led_green_off()
      led_red_on()
  end

  def color_white():
      led_blue_on()
      led_green_on()
      led_red_on()
  end

  def led_off():
      led_blue_off()
      led_green_off()
      led_red_off()
  end

  # COLOR FOR STATES
  thread Thread_Lights():
      while(True):
          # Stopping
          if (STATE == 1):
              color_red()
              sleep(0.5)
              led_off()
          # Stopped
          elif (STATE == 2):
              color_red()
          # Resetting
          # elif (STATE == 3):
          #     color_white()
          #     sleep(0.5)
          #     led_off()
          # Idle
          elif (AMR_Charging):
              color_white()
          # Starting
          # elif (STATE == 5):
          #     color_lightblue()
          #     sleep(0.5)
          #     led_off()
          # Execute
          # elif (STATE == 6):
          #     color_lightblue()
          # Completing
          # elif (STATE == 7):
          #     color_green()
          #     sleep(0.5)
          #     led_off()
          # # Complete
          # elif (STATE == 8):
          #     color_green()
          # Holding
          elif (STATE == 9):
              color_red()
              sleep(0.5)
              led_off()
          # Held
          elif (STATE == 10):
              color_red()
          # Unholding
          elif (STATE == 11):
              color_yellow()
              sleep(0.5)
              led_off()
          # Suspending
          elif (STATE == 12):
              color_blue()
              sleep(0.5)
              led_off()
          # Suspended
          elif (STATE == 13):
              color_blue()
          # Unsuspending
          elif (STATE == 14):
              color_yellow()
              sleep(0.5)
              led_off()
          # Aborting
          elif (STATE == 15):
              color_red()
              sleep(0.5)
              led_off()
          # Aborted
          elif (STATE == 16):
              color_red()
          # Clearing
          elif (STATE == 17):
              color_yellow()
              sleep(0.5)
              led_off()
          else:
              color_lightblue()
          end
          sleep(0.5)
      end
  end

  thread_lights_handler = run Thread_Lights()
  $ 10 "Script: SCRIPT Transitions V8.0.script"
  #*****************************************************
  # customer          :   INTERNAL
  # project name      :
  #****************************************************
  # controller        :   UR
  # software          :   5.13
  #****************************************************
  # author            :   P. Koehnke
  # Copyright (c)     :   United Robotics Group
  #                       An der Riede 2
  #                       28816 Stuhr
  #                       Germany
  #****************************************************
  # description       :   transition between workareas
  # version:      	:   1.2
  # created           :   28.02.2024
  # updated           :
  #****************************************************
  # modifications     :
  #
  # date              :
  # name              :
  # reason            :
  #****************************************************

  ######################### further development #########################
  #   - that the robot can switch the configuration, if necessary
  #   - introduction of structs
  #######################################################################

  ######################### to be adjusted #########################

  local WORKAREA_1 = [-0.280,-0.680,-0.001, 0.280, 0.100, 1.000]    # workarea 1 (platform)
  local WORKAREA_2 = [-1.000,-1.000,-1.000,-0.280, 0.100, 1.000]    # workarea 2 (front right)
  local WORKAREA_3 = [-1.000, 0.100,-1.000, 0.000, 1.000, 1.000]    # workarea 3 (back right)
  local WORKAREA_4 = [ 0.000, 0.100,-1.000, 1.000, 1.000, 1.000]    # workarea 4 (back left)
  local WORKAREA_5 = [ 0.280,-1.000,-1.000, 1.000, 0.100, 1.000]    # workarea 5 (front left)
  local WORKAREA_6 = [-0.280,-1.000,-1.000, 0.280,-0.680, 1.000]    # workarea 6 (front front)
  local WORKAREA_7 = [0,0,0,0,0,0]    # reserved
  local WORKAREA_8 = [0,0,0,0,0,0]    # reserved
  local WORKAREA_9 = [0,0,0,0,0,0]    # reserved
  local WORKAREA_10 = [0,0,0,0,0,0]   # reserved

  local PSE_WA_1 = p[ 0.000,-0.450, 0.300, 0.000, 0.000, 0.000]
  local PSE_WA_2 = p[-0.300,-0.300, 0.300, 0.000, 0.000, d2r(-90)]
  local PSE_WA_3 = p[-0.300, 0.300, 0.300, 0.000, 0.000, d2r(-135)]
  local PSE_WA_4 = p[ 0.300, 0.300, 0.300, 0.000, 0.000, d2r(135)]
  local PSE_WA_5 = p[ 0.300,-0.300, 0.300, 0.000, 0.000, d2r(90)]
  local PSE_WA_6 = p[ 0.000,-0.600, 0.300, 0.000, 0.000, 0.000]       # reserved
  local PSE_WA_7 = p[ 0.000, 0.000, 0.000, 0.000, 0.000, 0.000]       # reserved
  local PSE_WA_8 = p[ 0.000, 0.000, 0.000, 0.000, 0.000, 0.000]       # reserved
  local PSE_WA_9 = p[ 0.000, 0.000, 0.000, 0.000, 0.000, 0.000]       # reserved
  local PSE_WA_10 = p[ 0.000, 0.000, 0.000, 0.000, 0.000, 0.000]      # reserved

  global JNT_HOME = [-1.23163,-1.29627,-1.86552,-1.55102, 1.57761, 1.910]
  local JNT_STANDARD_C1 = [ 1.57,-1.57, 1.57,-1.57,-1.57,0]
  local JNT_STANDARD_C2 = [-1.57,-1.57,-1.57,-1.57, 1.57,0]
  local ANGLE_MIN_DEG = -110
  local ANGLE_MAX_DEG = 110
  local DISTANCE_TO_CLEARANCE = 0.300
  local RADIUS_HELPER_POSES = 0.300
  local RADIUS_TRANSITION_POSES = 0.400
  local workareas = [WORKAREA_1, WORKAREA_2, WORKAREA_3, WORKAREA_4, WORKAREA_5, WORKAREA_6, WORKAREA_7, WORKAREA_8, WORKAREA_9, WORKAREA_10]
  local poses = [PSE_WA_1, PSE_WA_2, PSE_WA_3, PSE_WA_4, PSE_WA_5, PSE_WA_6, PSE_WA_7, PSE_WA_8, PSE_WA_9, PSE_WA_10]

  ######################### end of adjustment #########################

  local pi = 3.14159265
  local axis_config_current = 0
  local axis_config_new = 0
  local workarea_current = 0
  local workarea_new = 0
  global reverse_rotation = False

  def create_translation_vector(x = 0.0, y = 0.0, z = 0.0):
      return struct(x = x, y = y, z = z)
  end

  def create_orientation_vector(rx = 0.0, ry = 0.0, rz = 0.0):
      return struct(rx = rx, ry = ry, rz = rz)
  end

  def create_transition_pose():
      return struct(crt = p[0,0,0,0,0,0], jnt = [0,0,0,0,0,0], q = [0,0,0,0,0,0], translation = create_translation_vector(), orientation = create_orientation_vector())
  end

  def compose_pose(translation = create_translation_vector(), orientation = create_orientation_vector()):
      return p[translation.x, translation.y, translation.z, orientation.rx, orientation.ry, orientation.rz]
  end

  local pose_start = create_transition_pose()
  local pose_help = create_transition_pose()
  local pose_target = create_transition_pose()
  local pose = create_transition_pose()

  def init_home_by_cartesian_pose(pose):
      # check given pose for reachability for the corresponding axis config
      local pose_home = pose_trans(pose, pose_inv(get_tcp_offset()))

      if check_current_axis_config() == 1:
          if get_inverse_kin_has_solution(pose_home, qnear=JNT_STANDARD_C1, tcp=p[0,0,0,0,0,0]):
              JNT_HOME = get_inverse_kin(pose_home, qnear=JNT_STANDARD_C1, tcp=p[0,0,0,0,0,0])
          end
      elif check_current_axis_config() == 2:
          if get_inverse_kin_has_solution(pose_home, qnear=JNT_STANDARD_C2, tcp=p[0,0,0,0,0,0]):
              JNT_HOME = get_inverse_kin(pose_home, qnear=JNT_STANDARD_C2, tcp=p[0,0,0,0,0,0])
          end
      end
  end

  def get_tool_free_pose(pose_ref=p[0,0,0,0,0,0], dir=[0,0,0], move_in_base_frame=False):
      # get a recovery pose
      # dir is providing the direction and distance in X, Y and Z
      # if 'move_in_base_frame' is set, dir will be interpreted as absolute values for a movement in base frame

      local pose_target = pose_ref
      local i = 0

      if pose_ref == p[0,0,0,0,0,0]:
          pose_target = get_actual_tcp_pose()
      end

      if (move_in_base_frame):
          while (i<3):
              # move only,
              # if the demanded position is bigger than zero and the current position is below the demanded one or
              # if the demanded position is smaller than zero and the current position is above the demanded one
              if ((dir[i]>0 and pose_target[i]<dir[i]) or (dir[i]<0 and pose_target[i]>dir[i])):
                  pose_target[i] = dir[i]
              end
              i = i + 1
          end
      else:
          pose_target = pose_trans(pose_ref, p[dir[0], dir[1], dir[2], 0, 0, 0])
      end

      return pose_target
  end

  def check_workarea(reference_pose):
      # the actual TCP position is compared to predefined areas (cubic) to determine in which area the robot arm is
      # a workarea is defined as a list of coordinates, where the first 3 values are X, Y, and Z with the smallest values and
      # the next 3 values specify X, Y and Z for the biggest values
      local data_size = size(workareas)
      local i = 0
      local size_workarea = p[0,0,0,0,0,0]
      local pose_workarea = p[0,0,0,0,0,0]

      while (i < data_size[0]):
          pose_workarea = pose_trans(inv(p[workareas[i, 0], workareas[i, 1], workareas[i, 2], 0, 0, 0]), reference_pose)
          size_workarea = pose_sub(p[workareas[i, 3], workareas[i, 4], workareas[i, 5], 0, 0, 0], p[workareas[i, 0], workareas[i, 1], workareas[i, 2], 0, 0, 0])
          if  ((pose_workarea[0]>0 and pose_workarea[0]<size_workarea[0]) and
              (pose_workarea[1]>0 and pose_workarea[1]<size_workarea[1]) and
              (pose_workarea[2]>0 and pose_workarea[2]<size_workarea[2])):
              return i + 1
          end
          i = i + 1
      end

      return 0
  end

  def check_current_axis_config():
      # function determnines, if the arm is oriented in one or the other configuration.
      # it means, that the ellbow joint is flipped and so are the wrist joints.

      local jnt_current = get_actual_joint_positions()

      # ellbow has positiv angle
      if (jnt_current[2]> 0):
          return 1
      # ellbow has negativ angle
      elif (jnt_current[2]< 0):
          return 2
      # angle is 0
      else:
          return 0
      end
  end

  def switch_axis_config(axis_config):
      # function to switch betwwen the axis configuration 1 and 2.

      if (axis_config == 1):
          return 2
      elif (axis_config ==2):
          return 1
      end
  end

  def get_joint_pose(pose, qnear):
      if get_inverse_kin_has_solution(pose, qnear=qnear):
          return get_inverse_kin(pose, qnear=qnear)
      else:
          popup("no solution found for the transition pose", blocking= True)
          return [0,0,0,0,0,0]
      end
  end

  def get_transition_pose_by_workarea(workarea):
      # get the correspondig pose from the list of poses

      pose.crt = poses[workarea-1]
      pose.q = set_q_near()
      pose.jnt = get_joint_pose(pose.crt, pose.q)

      return pose
  end

  def get_transition_pose_by_reference_pose(reference_pose, radius, keep_rxry=False):

      if reference_pose == p[0,0,0,0,0,0]:
          pose.jnt = JNT_HOME
          pose.q = JNT_HOME
          pose.crt = get_forward_kin(pose.jnt)
          if keep_rxry:
              pose.orientation = get_transition_orientation(pose.crt, keep_rxry)
              pose.crt = compose_pose(struct(x=pose.crt[0], y=pose.crt[1], z=pose.crt[2]), pose.orientation)
              pose.q = set_q_near(joints=[1,1,1,0,0,0])
              pose.jnt = get_joint_pose(pose.crt, pose.q)
          end
      else:
          pose.translation = get_transition_translation_by_radius(get_angle_to_base(reference_pose), radius)
          pose.orientation = get_transition_orientation(reference_pose, keep_rxry)
          pose.crt = compose_pose(pose.translation, pose.orientation)
          if keep_rxry:
              pose.q = set_q_near(joints=[1,1,1,0,0,0])
          else:
              pose.q = set_q_near(joints=[0,0,0,1,1,1])
          end
          pose.q[0] = adjust_axis_rotation(pose)
          pose.jnt = get_joint_pose(pose.crt, pose.q)
      end

      return pose
  end

  def get_rounded_mm(value):
      if (value < 0):
          return ceil(value*1000)
      elif (value >= 0):
          return floor(value*1000)
      end
  end

  def get_angle_to_base(pose):
      # get the angle relative to the base frame
      local pose_x_mm = 0
      local pose_y_mm = 0
      local angle = 0

      pose_x_mm = get_rounded_mm(pose[0])
      pose_y_mm = get_rounded_mm(pose[1])

      if (pose_x_mm == 0 and pose_y_mm < 0):
          angle = 0
      elif (pose_x_mm == 0 and pose_y_mm > 0):
          angle = pi
      elif (pose_x_mm < 0 and pose_y_mm == 0):
          angle = -pi/2
      elif (pose_x_mm > 0 and pose_y_mm == 0):
          angle = pi/2
      else:
          angle = atan2(pose[0], pose[1])
          if (-pi < angle) and (angle < 0):
              angle = - angle - pi
          elif (0 < angle) and (angle < pi):
              angle = - angle + pi
          end
      end
      return angle
  end

  def set_q_near(joints=[0,0,0,1,1,1], axis_config=check_current_axis_config()):
      local i = 0
      local jnt_current = get_actual_joint_positions()

      while i < 6:
          if joints[i] != 0:
              if axis_config == 1:
                  pose.q[i] = JNT_STANDARD_C1[i]
              elif axis_config == 2:
                  pose.q[i] = JNT_STANDARD_C2[i]
              else:
                  pose.q[i] = jnt_current[i]
              end
          else:
              pose.q[i] = jnt_current[i]
          end
          i = i + 1
      end
      return pose.q
  end

  def adjust_axis_rotation(pose):
      local angle = get_angle_to_base(pose.crt)

      if (0 > angle) and (angle > d2r(ANGLE_MIN_DEG)):
          if (pose.jnt[0] > JNT_HOME[0]):
              # calculated axis angle is in the wrong value range
              pose.q = set_q_near(joints=[1,0,0,0,0,0])
              reverse_rotation = True
          end
      elif (0 < angle) and (angle < d2r(ANGLE_MAX_DEG)):
          if (pose.jnt[0] < JNT_HOME[0]):
              pose.q = set_q_near(joints=[1,0,0,0,0,0])
              reverse_rotation = True
          end
      elif (pose.jnt[0] < -2 * pi):
          pose.q = set_q_near(joints=[1,0,0,0,0,0])
          reverse_rotation = True
      elif (pose.jnt[0] > 2 * pi):
          pose.q = set_q_near(joints=[1,0,0,0,0,0])
          reverse_rotation = True
      end
      return pose.q[0]
  end

  def get_transition_orientation(pose_ref, keep_rxry=False):
      # define the orientation of the transition poses
      local pose_current = get_actual_tcp_pose()
      local rpy_current = [0,0,0]
      local rotvec_new = [0,0,0]

      if keep_rxry:
          # use orientation of the given pose
          rpy_current = rotvec2rpy([pose_current[3], pose_current[4], pose_current[5]])
          rotvec_new = rpy2rotvec([rpy_current[0], rpy_current[1], get_angle_to_base(pose_ref) + get_locked_yaw()])
      else:
          # use orientation of defined workarea poses
          rpy_current = rotvec2rpy([pose_ref[3], pose_ref[4], pose_ref[5]])
          rotvec_new = rpy2rotvec([0, 0, rpy_current[2]])
      end
      return create_orientation_vector(rx = rotvec_new[0], ry = rotvec_new[1], rz = rotvec_new[2])
  end

  def get_transition_translation_by_radius(angle, radius):
      # calculate x,y by a radius and z by defined clearance
      return create_translation_vector(x = radius * cos(angle-pi/2), y = radius * sin(angle-pi/2), z = DISTANCE_TO_CLEARANCE)
  end

  def adjust_transition_poses(pose_identifier, keep_rxry=False):
      # adjust the orientation of the transition poses by determining the the current orientation

      local pose_current = get_actual_tcp_pose()
      local jnt_current = get_actual_joint_positions()
      local rpy_current = rotvec2rpy([pose_current[3],pose_current[4],pose_current[5]])
      local rotvec_new = [0,0,0]

      if (pose_identifier == "start"):
          pose = pose_start
      elif (pose_identifier == "target"):
          pose = pose_target
          pose.q[0] = adjust_axis_rotation(pose)
      elif (pose_identifier == "helper"):
          pose = pose_help
      end

      if keep_rxry:
          rotvec_new = rpy2rotvec([rpy_current[0], rpy_current[1], pose.angle_to_base + get_locked_yaw()])
          pose.crt = p[pose.crt[0], pose.crt[1], pose.crt[2], rotvec_new[0], rotvec_new[1], rotvec_new[2]]
          # adjust preferred joint angles ot the current ones
          pose.q[3] = jnt_current[3]
          pose.q[4] = jnt_current[4]
          pose.q[5] = jnt_current[5]
      end

      if get_inverse_kin_has_solution(pose.crt, qnear=pose.q) and is_within_safety_limits(pose.crt):
          pose.jnt = get_inverse_kin(pose.crt, qnear=pose.q)
      else:
          popup(str_cat("no solution for ", pose_identifier), error=True, blocking=False)
          pose.jnt = [0,0,0,0,0,0]
      end
      return pose.jnt
  end

  def get_locked_yaw():
      local pose_current = get_actual_tcp_pose()
      local rpy_current = rotvec2rpy([pose_current[3],pose_current[4],pose_current[5]])
      # local rotvec_new = rpy2rotvec([rpy_current[0], rpy_current[1], get_angle_to_base(pose_current)])
      local rotvec_new = rpy2rotvec([0, 0, get_angle_to_base(pose_current)])
      local pose_reference = p[pose_current[0], pose_current[1], pose_current[2], rotvec_new[0], rotvec_new[1], rotvec_new[2]]
      local pose_to_reference = pose_trans(pose_inv(pose_reference), pose_current)

      return pose_to_reference[5]
  end

  def get_helper_angle():
      local angle_start = get_angle_to_base(pose_start.crt)
      local angle_target = get_angle_to_base(pose_target.crt)
      local angle_help = (angle_start + angle_target) / 2

      if reverse_rotation and
          ((angle_start < 0 and
          angle_target < 0) or
          (angle_start > 0 and
          angle_target > 0)):
              angle_help = flip_angle(angle_help)
      elif (angle_start < 0 and
          angle_start < d2r(ANGLE_MIN_DEG)) and
          (angle_target > 0 and
          angle_target > d2r(ANGLE_MAX_DEG)):
              angle_help = flip_angle(angle_help)
      elif (angle_start > 0 and
          angle_start > d2r(ANGLE_MAX_DEG)) and
          (angle_target < 0 and
          angle_target < d2r(ANGLE_MIN_DEG)):
              angle_help = flip_angle(angle_help)
      end
      return angle_help
  end

  def flip_angle(angle):
      # flips the given angle 180 degree around
      if (angle < 0):
          return angle + pi
      elif (angle > 0):
          return angle - pi
      end
  end

